          MoveJ speed 100 deg/s, acceleration 80 deg/s^2 (useActiveTCP=true) feature=FRM_Reference
            Waypoint Variable (Variable): motionParameters(blendRadius=0.02); variable=PSE_A
        MoveL speed 400 mm/s, acceleration 500 mm/s^2 (useActiveTCP=true) feature=FRM_Reference
          Waypoint Variable (Variable): motionParameters(jointSpeed=1.047198 jointAcceleration=1.396263 cartesianSpeed=0.09 cartesianAcceleration=0.05); variable=PSE_T
          'ADD OPEN GRIPPER'
          URCap Gripper (Robotiq_Grippers, Robotiq Inc.) dataModel(position=78.82352941176471, force=11.0, speed=0.0, positionInDouble=78.82352941176471, forceInDouble=11.0, speedInDouble=0.0, slaveIds=[9], blocking=true)
          Waypoint Variable (Variable): motionParameters(jointSpeed=1.047198 jointAcceleration=1.396263 cartesianSpeed=0.09 cartesianAcceleration=0.05); variable=PSE_T_H
          URCap Gripper (Robotiq_Grippers, Robotiq Inc.) dataModel(position=24.705882352941178, force=11.0, speed=0.0, positionInDouble=24.705882352941178, forceInDouble=11.0, speedInDouble=0.0, slaveIds=[9], blocking=true)
          Waypoint Variable (Variable): variable=PSE_R
    Case (caseValue=7)
      Folder Load [hidden by the author, left out]
    Case (caseValue=8)
      Folder Unload [hidden by the author, left out]
    Case (caseValue=11)
      Folder Place without opening gripper
        Action_Info := "place object without gripper opening"
        SuppressedNode
          Script: do_transition(pose_trans(FRM_Reference, PSE_T), keep_rxry=OBJ_Picked)
        Script: movel(FRM_Container_S, a=0.025, v=0.015, r=0.00001)
        Folder EXTT
          Switch expression=JIG
            Case (caseValue=1)
              Folder 3FG
                If OBJ_Picked
                  Set DigitalOutput pin=GRP_3F_Open; digitalValue=1
        If PSE_A_H≠PSE_Z
          If JNT_Q≠JNT_Z
            Script: movej(get_inverse_kin(pose_trans(FRM_Reference, PSE_A_H), qnear=JNT_Q), r=0.050)
          Else 
            Script: movej(pose_trans(FRM_Reference, PSE_A_H), r=0.050)
        If PSE_A≠PSE_Z
          If JNT_Q≠JNT_Z
            Script: movej(get_inverse_kin(pose_trans(FRM_Reference, PSE_A), qnear=JNT_Q), r=0.020)
          Else 
            Script: movej(pose_trans(FRM_Reference, PSE_A), r=0.020)
        MoveL speed 400 mm/s, acceleration 500 mm/s^2 (useActiveTCP=true) feature=FRM_Reference
          If PSE_T_H≠PSE_Z
            Waypoint Variable (Variable): motionParameters(blendRadius=0.01); variable=PSE_T_H
          Waypoint Variable (Variable): motionParameters(jointSpeed=1.047198 jointAcceleration=1.396263 cartesianSpeed=0.09 cartesianAcceleration=0.05); variable=PSE_T
            Until TOOL_CONTACT_DETECTION (allowActions=false retraction=NONE decelerationAcceleration=0.5 decelerationAngularAcceleration=34.906585)
          Force Frame feature=FRM_Reference; selection=[1, 1, 1, 0, 0, 0]; wrench=[0, 0, 0, 0, 0, 0]; limitsForce=[0.1, 0.1, 0.01, 1.047198, 1.047198, 1.047198]; limitsMotion=[0.1, 0.1, 0.1, 0.349066, 0.349066, 0.349066]
            Waypoint Variable (Variable): motionParameters(jointSpeed=1.047198 jointAcceleration=1.396263 cartesianSpeed=0.07 cartesianAcceleration=0.04); variable=PSE_T
          Folder EXTT
            Switch expression=JIG
              Case (caseValue=1)
                Folder 3FG
                  If OBJ_Picked
                    Set DigitalOutput pin=GRP_3F_Open; digitalValue=0
                    Wait Sleep waitTime=0.2
          Folder EOAT
            ''
    Case (caseValue=12)
      Folder Decap
        Action_Info := "decapping"
        Set DigitalOutput pin=GRP_3F_Enable; digitalValue=1
        Set DigitalOutput pin=GRP_3F_Decap; digitalValue=1
        Force Simple feature=Joint_6_name; selection=[0, 0, 1, 0, 0, 0]; wrench=[0, 0, 5, 0, 0, 0]; limitsForce=[0.15, 0.15, 0.15, 1.047198, 1.047198, 1.047198]; limitsMotion=[0.1, 0.1, 0.1, 0.349066, 0.349066, 0.349066]
          Script: check_decapping(offset=0.015, timeout=5, abort=CMD_Hold)
        Set DigitalOutput pin=GRP_3F_Decap; digitalValue=0
        Set DigitalOutput pin=GRP_3F_Enable; digitalValue=0
        MoveL speed 150 mm/s, acceleration 800 mm/s^2 (useActiveTCP=true) feature=FRM_Reference
          Waypoint Variable (Variable): variable=PSE_R
    Case (caseValue=13)
      Timer (action=Reset) variable(name=TMR_Barcode)
      Folder Read [hidden by the author, left out]
    Case (caseValue=15)
      Folder Detect
        Action_Info := "detect"
    Case (caseValue=30)
      Folder Shake
        Action_Info := "shake"
        Script: do_transition(pose_trans(FRM_Reference, PSE_T), keep_rxry=OBJ_Picked)
        If PSE_A_H≠PSE_Z
          If JNT_Q≠JNT_Z
            Script: movej(get_inverse_kin(pose_trans(FRM_Reference, PSE_A_H), qnear=JNT_Q), r=0.050)
          Else 
            Script: movej(pose_trans(FRM_Reference, PSE_A_H), r=0.050)
        If PSE_A≠PSE_Z
          If JNT_Q≠JNT_Z
            Script: movej(get_inverse_kin(pose_trans(FRM_Reference, PSE_A), qnear=JNT_Q), r=0.020)
          Else 
            Script: movej(pose_trans(FRM_Reference, PSE_A), r=0.020)
        MoveL speed 400 mm/s, acceleration 500 mm/s^2 (useActiveTCP=true) feature=FRM_Reference
          If PSE_T_H≠PSE_Z
            Waypoint Variable (Variable): motionParameters(blendRadius=0.01); variable=PSE_T_H
          Waypoint Variable (Variable): motionParameters(jointSpeed=1.047198 jointAcceleration=1.396263 cartesianSpeed=0.12 cartesianAcceleration=0.08); variable=PSE_T
          Folder EXTT
            ''
            MoveJ speed 60 deg/s, acceleration 80 deg/s^2 (useActiveTCP=true) feature=Base
              Waypoint Waypoint_6: TCP in base x=8.801 y=-547.927 z=402.697 mm, rx=-0.5899 ry=-0.0072 rz=-0.0613 rad; joints [-69.01, -76.872, -104.694, -56.634, 78.043, -158.781] deg; TCP offset x=0 y=0 z=161 mm, rx=3.1415 ry=0 rz=0 rad
            MoveJ speed 60 deg/s, acceleration 80 deg/s^2 (useActiveTCP=true) feature=Base
              Waypoint Waypoint_18: TCP in base x=-178.372 y=-433.927 z=368.082 mm, rx=-0.0866 ry=0.7047 rz=-0.0079 rad; joints [-72.502, -76.524, -102.817, -99.71, 50.308, -158.785] deg
            MoveJ speed 60 deg/s, acceleration 80 deg/s^2 (useActiveTCP=true) feature=Base
              Waypoint Waypoint_12: TCP in base x=8.801 y=-547.927 z=402.697 mm, rx=-0.5899 ry=-0.0072 rz=-0.0613 rad; joints [-69.01, -76.872, -104.694, -56.634, 78.043, -158.781] deg
            MoveJ speed 60 deg/s, acceleration 80 deg/s^2 (useActiveTCP=true) feature=Base
              Waypoint Waypoint_19: TCP in base x=-178.372 y=-433.927 z=368.082 mm, rx=-0.0866 ry=0.7047 rz=-0.0079 rad; joints [-72.502, -76.524, -102.817, -99.71, 50.308, -158.785] deg
          If PSE_R_H≠PSE_Z
            Waypoint Variable (Variable): motionParameters(blendRadius=0.01); variable=PSE_R
            Waypoint Variable (Variable): variable=PSE_R_H
          Else 
            Waypoint Variable (Variable): variable=PSE_R
    Case (caseValue=31)
      Action_Info := "Pick_Vial"
      Folder Pick_Vial
        URCap Gripper (Robotiq_Grippers, Robotiq Inc.) dataModel(position=0.0, force=27.84313725490196, speed=32.15686274509804, positionInDouble=0.0, forceInDouble=27.84313725490196, speedInDouble=32.15686274509804, slaveIds=[9], blocking=true)
        MoveJ speed 60 deg/s, acceleration 80 deg/s^2 (useActiveTCP=true) feature=Base
          Waypoint Vial_above: motionParameters(jointSpeed=0.436332 jointAcceleration=0.523599 cartesianSpeed=0.25 cartesianAcceleration=1.2 blendRadius=0.05); TCP in base x=17.106 y=-652.093 z=184.921 mm, rx=0 ry=0 rz=1.5641 rad; joints [-76.636, -112.403, -84.029, -73.556, 90.141, -256.27] deg
        MoveL speed 250 mm/s, acceleration 1200 mm/s^2 (useActiveTCP=true) feature=Base
          Waypoint Vial_pick_point: motionParameters(jointSpeed=1.047198 jointAcceleration=1.396263 cartesianSpeed=0.1 cartesianAcceleration=0.5); TCP in base x=17.106 y=-648.923 z=93.308 mm, rx=0 ry=0 rz=1.5641 rad; joints [-76.583, -116.742, -92.083, -61.164, 90.132, -256.177] deg
        URCap Gripper (Robotiq_Grippers, Robotiq Inc.) dataModel(position=100.0, force=32.94117647058823, speed=27.84313725490196, positionInDouble=100.0, forceInDouble=32.94117647058823, speedInDouble=27.84313725490196, slaveIds=[9], blocking=true)
        MoveL speed 250 mm/s, acceleration 1200 mm/s^2 (useActiveTCP=true) feature=Base
          Waypoint Waypoint_20: motionParameters(jointSpeed=1.047198 jointAcceleration=1.396263 cartesianSpeed=0.1 cartesianAcceleration=0.5 blendRadius=0.05); TCP in base x=19.228 y=-648.67 z=184.921 mm, rx=0 ry=0 rz=0.0241 rad; joints [-76.382, -111.96, -84.66, -73.372, 90.146, -167.779] deg
        SafeHome (positionOptionType=SPEED_AND_ACCELERATION speed=1.047198 acceleration=1.396263 nextMotionTime=2)
    Case (caseValue=32)
      decap := False
      Folder decap_Vial
        Set DigitalOutput pin=digital_out[5]; digitalValue=1
        MoveJ speed 60 deg/s, acceleration 80 deg/s^2 (useActiveTCP=true) feature=Base
          Waypoint Waypoint_33: motionParameters(jointSpeed=0.436332 jointAcceleration=0.523599 cartesianSpeed=0.25 cartesianAcceleration=1.2 blendRadius=0); TCP in base x=-32.362 y=-348.336 z=391.476 mm, rx=0 ry=0 rz=-0.0047 rad; joints [-72.819, -68.266, -97.918, -103.808, 90.124, -162.602] deg
        MoveL speed 250 mm/s, acceleration 1200 mm/s^2 (useActiveTCP=true) feature=Base
          Waypoint Vial_3FG_place: motionParameters(jointSpeed=1.047198 jointAcceleration=1.396263 cartesianSpeed=0.1 cartesianAcceleration=0.5); TCP in base x=-31.859 y=-349.403 z=145.301 mm, rx=0 ry=0 rz=0 rad; joints [-72.903, -71.756, -132.514, -65.722, 90.129, -162.805] deg
        Set DigitalOutput pin=digital_out[5]; digitalValue=0
        Wait Sleep waitTime=0.5
        MoveL speed 250 mm/s, acceleration 1200 mm/s^2 (useActiveTCP=true) feature=Base
          Waypoint Waypoint_34: motionParameters(jointSpeed=1.047198 jointAcceleration=1.396263 cartesianSpeed=0.1 cartesianAcceleration=0.5 blendRadius=0.05); TCP in base x=-32.362 y=-348.336 z=391.476 mm, rx=0 ry=0 rz=-0.0047 rad; joints [-72.819, -68.266, -97.918, -103.808, 90.124, -162.602] deg
        MoveJ speed 60 deg/s, acceleration 80 deg/s^2 (useActiveTCP=true) feature=Base
          Waypoint cap_dump: motionParameters(jointSpeed=0.436332 jointAcceleration=0.523599 cartesianSpeed=0.25 cartesianAcceleration=1.2); TCP in base x=-139.169 y=-420.164 z=146.096 mm, rx=0 ry=0 rz=0 rad; joints [-90.79, -86.479, -121, -62.513, 90.12, -180.712] deg
        URCap Gripper (Robotiq_Grippers, Robotiq Inc.) dataModel(position=0.0, force=100.0, speed=100.0, positionInDouble=0.0, forceInDouble=100.0, speedInDouble=100.0, slaveIds=[9], blocking=true)
        MoveJ speed 60 deg/s, acceleration 80 deg/s^2 (useActiveTCP=true) feature=Base
          Waypoint Waypoint_35: motionParameters(jointSpeed=0.436332 jointAcceleration=0.523599 cartesianSpeed=0.25 cartesianAcceleration=1.2 blendRadius=0.05); TCP in base x=-32.362 y=-348.336 z=391.476 mm, rx=0 ry=0 rz=-0.0047 rad; joints [-72.819, -68.266, -97.918, -103.808, 90.124, -162.602] deg
        MoveL speed 250 mm/s, acceleration 1200 mm/s^2 (useActiveTCP=true) feature=Base
          Waypoint Vial_3FG_place: motionParameters(jointSpeed=1.047198 jointAcceleration=1.396263 cartesianSpeed=0.1 cartesianAcceleration=0.5); TCP in base x=-31.859 y=-349.403 z=145.301 mm, rx=0 ry=0 rz=0 rad; joints [-72.903, -71.756, -132.514, -65.722, 90.129, -162.805] deg
        URCap Gripper (Robotiq_Grippers, Robotiq Inc.) dataModel(position=100.0, force=100.0, speed=80.0, positionInDouble=100.0, forceInDouble=100.0, speedInDouble=80.0, slaveIds=[9], blocking=true)
        SuppressedNode
          decap := True
        SuppressedNode
          Script: dynamic_upward_motion(0.015, 7)
        SuppressedNode
          MoveL speed 250 mm/s, acceleration 1200 mm/s^2 (useActiveTCP=true) feature=Joint_6_name
            MoveDirectionNode (selectedDirection=ZPlus toolParams=8.0E-4, 0.001) feature=Base
              Until DISTANCE (allowActions=false deceleration=3 distanceNodeType=STOP) Distance=0.01; motionParameters(blendRadius=0)
        SuppressedNode
          decap := False
        Folder Decap
          Action_Info := "decapping"
          Set DigitalOutput pin=GRP_3F_Enable; digitalValue=1
          Set DigitalOutput pin=GRP_3F_Decap; digitalValue=1
          Force Frame feature=Base; selection=[0, 0, 1, 0, 0, 0]; wrench=[0, 0, 1, 0, 0, 0]; limitsForce=[0.15, 0.15, 0.001, 1.047198, 1.047198, 1.047198]; limitsMotion=[0.1, 0.1, 0.1, 0.349066, 0.349066, 0.349066]
            Script: check_decapping(offset=0.015, timeout=10, abort=CMD_Hold)
          Set DigitalOutput pin=GRP_3F_Decap; digitalValue=0
          Set DigitalOutput pin=GRP_3F_Enable; digitalValue=0
          MoveL speed 250 mm/s, acceleration 1200 mm/s^2 (useActiveTCP=true) feature=Base
            Waypoint Waypoint_36: motionParameters(jointSpeed=1.047198 jointAcceleration=1.396263 cartesianSpeed=0.1 cartesianAcceleration=0.5 blendRadius=0.05); TCP in base x=-32.362 y=-348.336 z=391.476 mm, rx=0 ry=0 rz=-0.0047 rad; joints [-72.819, -68.266, -97.918, -103.808, 90.124, -162.602] deg
        MoveJ speed 60 deg/s, acceleration 80 deg/s^2 (useActiveTCP=true) feature=Base
          Waypoint cap_dump: motionParameters(jointSpeed=0.436332 jointAcceleration=0.523599 cartesianSpeed=0.25 cartesianAcceleration=1.2); TCP in base x=-139.169 y=-420.164 z=146.096 mm, rx=0 ry=0 rz=0 rad; joints [-90.79, -86.479, -121, -62.513, 90.12, -180.712] deg
        URCap Gripper (Robotiq_Grippers, Robotiq Inc.) dataModel(position=0.0, force=100.0, speed=80.0, positionInDouble=0.0, forceInDouble=100.0, speedInDouble=80.0, slaveIds=[9], blocking=true)
        MoveJ speed 60 deg/s, acceleration 80 deg/s^2 (useActiveTCP=true) feature=Base
          Waypoint Waypoint_37: motionParameters(jointSpeed=0.436332 jointAcceleration=0.523599 cartesianSpeed=0.25 cartesianAcceleration=1.2 blendRadius=0.036); TCP in base x=-32.362 y=-348.336 z=391.476 mm, rx=0 ry=0 rz=-0.0047 rad; joints [-72.819, -68.266, -97.918, -103.808, 90.124, -162.602] deg
    Case (caseValue=33)
      Folder Shake and liquid transfer
        MoveL speed 250 mm/s, acceleration 1200 mm/s^2 (useActiveTCP=true) feature=Base
          Waypoint Vial_liq_above: motionParameters(jointSpeed=1.047198 jointAcceleration=1.396263 cartesianSpeed=0.1 cartesianAcceleration=0.5); TCP in base x=-25.304 y=-338.759 z=426.628 mm, rx=-1.3159 ry=0.8 rz=-0.9283 rad; joints [-21.713, -86.8, -129.663, 45.096, -43.028, -184.708] deg
          Waypoint Vial_liq_pick_1: motionParameters(jointSpeed=1.047198 jointAcceleration=1.396263 cartesianSpeed=0.1 cartesianAcceleration=0.5); TCP in base x=-2.66 y=-335.985 z=159.39 mm, rx=-1.1505 ry=0.6732 rz=-1.0106 rad; joints [-20.975, -83.1, -137.831, -114.287, 46.064, -14.375] deg
          Waypoint Vial_liq_pick_2: motionParameters(jointSpeed=1.047198 jointAcceleration=1.396263 cartesianSpeed=0.1 cartesianAcceleration=0.5); TCP in base x=-41.402 y=-356.792 z=125.395 mm, rx=-1.1435 ry=0.6511 rz=-0.8787 rad; joints [-25.36, -82.348, -146.215, -101.788, 37.598, -24.648] deg
          URCap Gripper (Robotiq_Grippers, Robotiq Inc.) dataModel(position=100.0, force=27.84313725490196, speed=32.15686274509804, positionInDouble=100.0, forceInDouble=27.84313725490196, speedInDouble=32.15686274509804, slaveIds=[9], blocking=true)
          Wait Sleep waitTime=1
          Set DigitalOutput pin=digital_out[5]; digitalValue=1
          Wait Sleep waitTime=0.5
          Waypoint Vial_liq_above: motionParameters(jointSpeed=1.047198 jointAcceleration=1.396263 cartesianSpeed=0.05 cartesianAcceleration=0.3 blendRadius=0.05); TCP in base x=-25.304 y=-338.759 z=426.628 mm, rx=-1.3159 ry=0.8 rz=-0.9283 rad; joints [-21.713, -86.8, -129.663, 45.096, -43.028, -184.708] deg
        MoveL speed 250 mm/s, acceleration 1200 mm/s^2 (useActiveTCP=true) feature=Base
          Waypoint Liquid_midway: motionParameters(jointSpeed=1.047198 jointAcceleration=1.396263 cartesianSpeed=0.1 cartesianAcceleration=0.5 blendRadius=0); TCP in base x=57.575 y=-583.082 z=306.415 mm, rx=-1.3517 ry=0.1209 rz=-0.0969 rad; joints [-51.29, -97.606, -136.419, 36.185, 44.156, -168.768] deg
          Loop Counting (count=3) loopVariable(name=Loop_1)
            Waypoint shake_1: motionParameters(jointSpeed=1.047198 jointAcceleration=1.396263 cartesianSpeed=0.5 cartesianAcceleration=2); TCP in base x=57.575 y=-583.085 z=306.423 mm, rx=-1.361 ry=-0.1556 rz=-0.4381 rad; joints [-51.29, -97.606, -136.418, 36.185, 44.156, -145.5] deg
            Waypoint shake_2: motionParameters(jointSpeed=1.047198 jointAcceleration=1.396263 cartesianSpeed=0.5 cartesianAcceleration=2); TCP in base x=57.582 y=-583.091 z=306.44 mm, rx=-1.3088 ry=0.3685 rz=0.2149 rad; joints [-51.29, -97.606, -136.416, 36.185, 44.155, -190] deg
          Waypoint drop_above_1: motionParameters(jointSpeed=1.047198 jointAcceleration=1.396263 cartesianSpeed=0.1 cartesianAcceleration=0.5); TCP in base x=268.235 y=-467.784 z=226.22 mm, rx=-1.0278 ry=-0.4308 rz=1.0046 rad; joints [-53.609, -95.474, -138.959, 24.045, 105.829, -198.245] deg
          Waypoint drop_above_2: motionParameters(jointSpeed=1.047198 jointAcceleration=1.396263 cartesianSpeed=0.1 cartesianAcceleration=0.5); TCP in base x=219.042 y=-470.776 z=133.754 mm, rx=-0.313 ry=-0.3444 rz=1.5006 rad; joints [-60.743, -97.429, -119.175, -41.501, 111.324, -235.78] deg
          Waypoint liq_tran_1: motionParameters(jointSpeed=1.047198 jointAcceleration=1.396263 cartesianSpeed=0.05 cartesianAcceleration=0.5 blendRadius=0.008); TCP in base x=213.068 y=-469.567 z=100.231 mm, rx=0.2519 ry=0.2179 rz=1.5928 rad; joints [-44.631, -104.414, -106.819, -71.743, 78.886, -225.335] deg
          Wait Sleep waitTime=1
          Waypoint drop_above_2: motionParameters(jointSpeed=1.047198 jointAcceleration=1.396263 cartesianSpeed=0.1 cartesianAcceleration=0.5); TCP in base x=219.042 y=-470.776 z=133.754 mm, rx=-0.313 ry=-0.3444 rz=1.5006 rad; joints [-60.743, -97.429, -119.175, -41.501, 111.324, -235.78] deg
          Waypoint Waypoint_21: motionParameters(jointSpeed=1.047198 jointAcceleration=1.396263 cartesianSpeed=0.1 cartesianAcceleration=0.5); TCP in base x=187.119 y=-493.959 z=133.754 mm, rx=-0.313 ry=-0.3444 rz=1.5006 rad; joints [-65.422, -99.182, -116.519, -44.234, 112.218, -240.733] deg
          Waypoint liq_tran_2: motionParameters(jointSpeed=1.047198 jointAcceleration=1.396263 cartesianSpeed=0.05 cartesianAcceleration=0.5); TCP in base x=195.958 y=-493.023 z=100.231 mm, rx=0.1607 ry=0.1098 rz=1.5253 rad; joints [-50.52, -104.533, -106.862, -66.514, 83.832, -227.689] deg
          Wait Sleep waitTime=1
          Waypoint drop_above_2: motionParameters(jointSpeed=1.047198 jointAcceleration=1.396263 cartesianSpeed=0.1 cartesianAcceleration=0.5); TCP in base x=219.042 y=-470.776 z=133.754 mm, rx=-0.313 ry=-0.3444 rz=1.5006 rad; joints [-60.743, -97.429, -119.175, -41.501, 111.324, -235.78] deg
          Waypoint drop_above_1: motionParameters(jointSpeed=1.047198 jointAcceleration=1.396263 cartesianSpeed=0.1 cartesianAcceleration=0.5); TCP in base x=268.235 y=-467.784 z=226.22 mm, rx=-1.0278 ry=-0.4308 rz=1.0046 rad; joints [-53.609, -95.474, -138.959, 24.045, 105.829, -198.245] deg
          Waypoint Liquid_midway: motionParameters(jointSpeed=1.047198 jointAcceleration=1.396263 cartesianSpeed=0.1 cartesianAcceleration=0.5); TCP in base x=57.575 y=-583.082 z=306.415 mm, rx=-1.3517 ry=0.1209 rz=-0.0969 rad; joints [-51.29, -97.606, -136.419, 36.185, 44.156, -168.768] deg
        MoveL speed 250 mm/s, acceleration 1200 mm/s^2 (useActiveTCP=true) feature=Base
          Waypoint Vial_drop_above: motionParameters(jointSpeed=1.047198 jointAcceleration=1.396263 cartesianSpeed=0.1 cartesianAcceleration=0.5); TCP in base x=0.325 y=-648.57 z=221.894 mm, rx=-0.8735 ry=1.1659 rz=-1.4827 rad; joints [-60.601, -137.11, -52.92, -147.418, 45.283, -19.072] deg
          Waypoint Vial_liq_drop: motionParameters(jointSpeed=1.047198 jointAcceleration=1.396263 cartesianSpeed=0.1 cartesianAcceleration=0.5); TCP in base x=1.021 y=-647.66 z=92.916 mm, rx=-0.8348 ry=1.0819 rz=-1.5406 rad; joints [-60.917, -140.075, -64.676, -125.954, 46.582, -22.337] deg
          URCap Gripper (Robotiq_Grippers, Robotiq Inc.) dataModel(position=0.0, force=27.84313725490196, speed=32.15686274509804, positionInDouble=0.0, forceInDouble=27.84313725490196, speedInDouble=32.15686274509804, slaveIds=[9], blocking=true)
          Waypoint Vial_drop_above: motionParameters(jointSpeed=1.047198 jointAcceleration=1.396263 cartesianSpeed=0.1 cartesianAcceleration=0.5); TCP in base x=0.325 y=-648.57 z=221.894 mm, rx=-0.8735 ry=1.1659 rz=-1.4827 rad; joints [-60.601, -137.11, -52.92, -147.418, 45.283, -19.072] deg
    Case (caseValue=34)
      SafeHome (positionOptionType=SPEED_AND_ACCELERATION speed=1.047198 acceleration=1.396263 nextMotionTime=2)
      MoveJ speed 60 deg/s, acceleration 80 deg/s^2 (useActiveTCP=true) feature=Base
        Waypoint Waypoint_9: motionParameters(jointSpeed=0.436332 jointAcceleration=0.523599 cartesianSpeed=0.25 cartesianAcceleration=1.2); TCP in base x=206.301 y=-401.796 z=209.941 mm, rx=0 ry=0 rz=1.5608 rad; joints [-45.627, -84.145, -113.025, -72.821, 90.127, -225.014] deg
      MoveL speed 250 mm/s, acceleration 1200 mm/s^2 (useActiveTCP=true) feature=Base
        Waypoint Waypoint_10: motionParameters(jointSpeed=1.047198 jointAcceleration=1.396263 cartesianSpeed=0.1 cartesianAcceleration=0.5); TCP in base x=200.866 y=-400.818 z=105.073 mm, rx=0 ry=0 rz=1.5608 rad; joints [-46.083, -90.669, -123.933, -55.389, 90.105, -225.416] deg
      URCap Gripper (Robotiq_Grippers, Robotiq Inc.) dataModel(position=100.0, force=27.84313725490196, speed=32.15686274509804, positionInDouble=100.0, forceInDouble=27.84313725490196, speedInDouble=32.15686274509804, slaveIds=[9], blocking=true)
      Wait Sleep waitTime=1
      MoveL speed 250 mm/s, acceleration 1200 mm/s^2 (useActiveTCP=true) feature=Base
        Waypoint Waypoint_11: motionParameters(jointSpeed=1.047198 jointAcceleration=1.396263 cartesianSpeed=0.1 cartesianAcceleration=0.5 blendRadius=0.05); TCP in base x=200.866 y=-400.818 z=325.177 mm, rx=0 ry=0 rz=1.5608 rad; joints [-46.018, -81.306, -98.396, -90.289, 90.129, -225.47] deg
      MoveJ speed 60 deg/s, acceleration 80 deg/s^2 (useActiveTCP=true) feature=Base
        Waypoint Waypoint_7: motionParameters(jointSpeed=0.436332 jointAcceleration=0.523599 cartesianSpeed=0.25 cartesianAcceleration=1.2 blendRadius=0.05); TCP in base x=-615.829 y=233.809 z=300 mm, rx=0.0051 ry=0.0087 rz=-2.1118 rad; joints [-188.832, -110.936, -69.076, -89.912, 89.674, -157.919] deg
      MoveL speed 250 mm/s, acceleration 1200 mm/s^2 (useActiveTCP=true) feature=Base
        Waypoint Waypoint_8: motionParameters(jointSpeed=1.047198 jointAcceleration=1.396263 cartesianSpeed=0.1 cartesianAcceleration=0.5); TCP in base x=-615.829 y=233.809 z=13.91 mm, rx=0.0051 ry=0.0087 rz=-2.1118 rad; joints [-188.874, -123.68, -94.539, -51.707, 89.657, -157.833] deg
      URCap Gripper (Robotiq_Grippers, Robotiq Inc.) dataModel(position=0.0, force=27.84313725490196, speed=32.15686274509804, positionInDouble=0.0, forceInDouble=27.84313725490196, speedInDouble=32.15686274509804, slaveIds=[9], blocking=true)
      MoveJ speed 60 deg/s, acceleration 80 deg/s^2 (useActiveTCP=true) feature=Base
        Waypoint Waypoint_7: motionParameters(jointSpeed=0.436332 jointAcceleration=0.523599 cartesianSpeed=0.25 cartesianAcceleration=1.2); TCP in base x=-615.829 y=233.809 z=300 mm, rx=0.0051 ry=0.0087 rz=-2.1118 rad; joints [-188.832, -110.936, -69.076, -89.912, 89.674, -157.919] deg
      SafeHome (positionOptionType=SPEED_AND_ACCELERATION speed=1.047198 acceleration=1.396263 nextMotionTime=2)
      SuppressedNode
        Folder Decap
          Action_Info := "decapping"
          Set DigitalOutput pin=GRP_3F_Enable; digitalValue=1
          Set DigitalOutput pin=GRP_3F_Decap; digitalValue=1
          Force Frame feature=Base; selection=[0, 0, 1, 0, 0, 0]; wrench=[0, 0, 1, 0, 0, 0]; limitsForce=[0.15, 0.15, 0.001, 1.047198, 1.047198, 1.047198]; limitsMotion=[0.1, 0.1, 0.1, 0.349066, 0.349066, 0.349066]
            Script: check_decapping(offset=0.015, timeout=10, abort=CMD_Hold)
          Set DigitalOutput pin=GRP_3F_Decap; digitalValue=0
          Set DigitalOutput pin=GRP_3F_Enable; digitalValue=0
          MoveL speed 250 mm/s, acceleration 1200 mm/s^2 (useActiveTCP=true) feature=Base
            Waypoint Waypoint_5: motionParameters(jointSpeed=1.047198 jointAcceleration=1.396263 cartesianSpeed=0.1 cartesianAcceleration=0.5 blendRadius=0.05); TCP in base x=-31.859 y=-349.402 z=312.809 mm, rx=0 ry=0 rz=0 rad; joints [-72.832, -66.838, -110.376, -92.778, 90.139, -162.834] deg
          MoveJ speed 60 deg/s, acceleration 80 deg/s^2 (useActiveTCP=true) feature=Base
            Waypoint cap_dump: motionParameters(jointSpeed=0.436332 jointAcceleration=0.523599 cartesianSpeed=0.25 cartesianAcceleration=1.2); TCP in base x=-139.169 y=-420.164 z=146.096 mm, rx=0 ry=0 rz=0 rad; joints [-90.79, -86.479, -121, -62.513, 90.12, -180.712] deg
          URCap Gripper (Robotiq_Grippers, Robotiq Inc.) dataModel(position=0.0, force=100.0, speed=100.0, positionInDouble=0.0, forceInDouble=100.0, speedInDouble=100.0, slaveIds=[9], blocking=true)
          MoveJ speed 60 deg/s, acceleration 80 deg/s^2 (useActiveTCP=true) feature=Base
            Waypoint Waypoint_5: motionParameters(jointSpeed=0.436332 jointAcceleration=0.523599 cartesianSpeed=0.25 cartesianAcceleration=1.2 blendRadius=0.05); TCP in base x=-31.859 y=-349.402 z=312.809 mm, rx=0 ry=0 rz=0 rad; joints [-72.832, -66.838, -110.376, -92.778, 90.139, -162.834] deg
          Set DigitalOutput pin=digital_out[5]; digitalValue=1
    Case (caseValue=35)
      Folder Pick the powder container
        SuppressedNode
          MoveJ speed 60 deg/s, acceleration 80 deg/s^2 (useActiveTCP=true) feature=Base
            Waypoint Variable (Variable): variable(featureName=CAM_LM_Cont_S)
        URCap VISOR Robotic App (SensoPart VISOR Robotic, SensoPart Industriesensorik GmbH) dataModel(visorAppTemplate=1); state(isChildrenLocked=true)
          URCap Easy Pick Setup (SensoPart VISOR Robotic, SensoPart Industriesensorik GmbH) dataModel(visorId=0, visorSetJob=true, visorImageAcqSetup=2, visorDetector=1, visorOffsetSet=true, visorCalibSetNo=7, visorJobName=Container, visorImageAcqSource=2, visorSetupStatus=2, Pose(key=visorImageAcqPose, Position(key=posePosition, Length(key=X value=-0.51041 unit=M), Length(key=Y value=0.417301 unit=M), Length(key=Z value=0.464095 unit=M)), Rotation(key=poseRotation, Angle(key=RX value=0.000026 unit=RAD), Angle(key=RY value=-0.000024 unit=RAD), Angle(key=RZ value=-2.896187 unit=RAD))), Pose(key=visorGripPose, Position(key=posePosition, Length(key=X value=-0.52891 unit=M), Length(key=Y value=0.461593 unit=M), Length(key=Z value=-0.178186 unit=M)), Rotation(key=poseRotation, Angle(key=RX value=-0.279814 unit=RAD), Angle(key=RY value=2.118244 unit=RAD), Angle(key=RZ value=-2.110314 unit=RAD))), Feature(key=visorImageAcqFeature name=cont_img_pose)); state(isChildrenLocked=true)
          URCap Process (SensoPart VISOR Robotic, SensoPart Industriesensorik GmbH) dataModel(Variable(key=visorCounterVar, variable(name=easyPickCount, initializeExpression=0)), Variable(key=visorPartsFoundVar, variable(name=easyPickParts, initializeExpression=0))); state(isChildrenLocked=true)
            URCap Image Acquisition Pose (SensoPart VISOR Robotic, SensoPart Industriesensorik GmbH) state(isChildrenLocked=true)
            URCap Object Detected (SensoPart VISOR Robotic, SensoPart Industriesensorik GmbH) state(isChildrenLocked=true)
              Folder Open Gripper
                URCap Gripper (Robotiq_Grippers, Robotiq Inc.) dataModel(position=0.0, force=30.0, speed=40.0, positionInDouble=0.0, forceInDouble=30.0, speedInDouble=40.0, slaveIds=[9], blocking=true)
                MoveJ speed 60 deg/s, acceleration 80 deg/s^2 (useActiveTCP=true) feature=Base
                  Waypoint Waypoint_13: TCP in base x=-479.451 y=284.141 z=125.27 mm, rx=-0.2768 ry=2.0984 rz=-2.1213 rad; joints [-165.671, -112.009, -127.874, -95.426, 1.192, -23.029] deg
              URCap Approach Pose (SensoPart VISOR Robotic, SensoPart Industriesensorik GmbH) dataModel(visorOffsetZ=-50.0); state(isChildrenLocked=true)
              URCap Target Pose (SensoPart VISOR Robotic, SensoPart Industriesensorik GmbH) state(isChildrenLocked=true)
              Folder Close Gripper
                URCap Gripper (Robotiq_Grippers, Robotiq Inc.) dataModel(position=100.0, force=30.19607843137255, speed=40.0, positionInDouble=100.0, forceInDouble=30.19607843137255, speedInDouble=40.0, slaveIds=[9], blocking=true)
              URCap Exit Pose (SensoPart VISOR Robotic, SensoPart Industriesensorik GmbH) dataModel(visorOffsetZ=-50.0); state(isChildrenLocked=true)
            URCap No Object Detected (SensoPart VISOR Robotic, SensoPart Industriesensorik GmbH) dataModel(Variable(key=visorNoObjCountVar, variable(name=easyPickNoObj, initializeExpression=0)))
              Popup Message (haltProgram=false message=No Container detected inputType=Text)
        MoveJ speed 60 deg/s, acceleration 80 deg/s^2 (useActiveTCP=true) feature=Base
          SuppressedNode
            Waypoint Cont_midwa_1: motionParameters(jointSpeed=1.047198 jointAcceleration=1.396263 cartesianSpeed=0.25 cartesianAcceleration=1.2 blendRadius=0.01); TCP in base x=-462.252 y=294.856 z=204.322 mm, rx=-0.3472 ry=2.0343 rz=-2.0655 rad; joints [-166.773, -128.859, -129.893, 70.604, 5.32, -171.145] deg
          Waypoint Waypoint_70: motionParameters(jointSpeed=0.523599 jointAcceleration=0.698132 cartesianSpeed=0.25 cartesianAcceleration=1.2 blendRadius=0); TCP in base x=-472.821 y=292.44 z=207.418 mm, rx=-0.2598 ry=-2.0535 rz=2.0707 rad; joints [-170.164, -118.699, -96.461, -142.976, 25.725, -0.32] deg
          Waypoint Waypoint_2: motionParameters(jointSpeed=0.523599 jointAcceleration=0.872665 cartesianSpeed=0.25 cartesianAcceleration=1.2 blendRadius=0.05); TCP in base x=-312.961 y=-152.991 z=223.61 mm, rx=-0.7453 ry=-1.7139 rz=1.6733 rad; joints [-134.992, -125.122, -83.555, -151.463, 94.666, 2.49] deg
          Waypoint Waypoint_3: motionParameters(jointSpeed=0.523599 jointAcceleration=0.698132 cartesianSpeed=0.25 cartesianAcceleration=1.2 blendRadius=0.05); TCP in base x=-113.75 y=-390.11 z=317.307 mm, rx=-0.5194 ry=-0.8399 rz=1.7569 rad; joints [-108.345, -98.585, -86.606, -121.699, 124.957, 41.411] deg
        MoveL speed 250 mm/s, acceleration 1200 mm/s^2 (useActiveTCP=true) feature=Base
          Waypoint Waypoint_15: motionParameters(jointSpeed=1.047198 jointAcceleration=1.396263 cartesianSpeed=0.1 cartesianAcceleration=0.5 blendRadius=0.05); TCP in base x=29.144 y=-436.802 z=327.885 mm, rx=-0.5216 ry=-0.6236 rz=1.8627 rad; joints [-89.657, -89.204, -96.411, -97.086, 128.129, 64.023] deg
          Waypoint Waypoint_14: motionParameters(jointSpeed=1.047198 jointAcceleration=1.396263 cartesianSpeed=0.1 cartesianAcceleration=0.3); TCP in base x=68.712 y=-569.42 z=285.215 mm, rx=-0.6792 ry=-0.7121 rz=1.394 rad; joints [-90.137, -103.3, -96.148, -70.007, 141.633, 93.932] deg
          Waypoint Waypoint_4: motionParameters(jointSpeed=1.047198 jointAcceleration=1.396263 cartesianSpeed=0.05 cartesianAcceleration=0.3); TCP in base x=-47.22 y=-557.625 z=136.371 mm, rx=-0.6792 ry=-0.7121 rz=1.394 rad; joints [-101.643, -114.727, -100.71, -68.127, 140.302, 75.797] deg
        URCap Gripper (Robotiq_Grippers, Robotiq Inc.) dataModel(position=0.0, force=30.0, speed=40.0, positionInDouble=0.0, forceInDouble=30.0, speedInDouble=40.0, slaveIds=[9], blocking=true)
        MoveL speed 250 mm/s, acceleration 1200 mm/s^2 (useActiveTCP=true) feature=Base
          Waypoint Waypoint_25: motionParameters(jointSpeed=1.047198 jointAcceleration=1.396263 cartesianSpeed=0.1 cartesianAcceleration=0.3); TCP in base x=65.436 y=-569.388 z=287.821 mm, rx=-0.6792 ry=-0.7121 rz=1.394 rad; joints [-90.466, -103.248, -95.699, -70.925, 141.635, 93.398] deg
          Waypoint Waypoint_15: motionParameters(jointSpeed=1.047198 jointAcceleration=1.396263 cartesianSpeed=0.1 cartesianAcceleration=0.5 blendRadius=0.05); TCP in base x=29.144 y=-436.802 z=327.885 mm, rx=-0.5216 ry=-0.6236 rz=1.8627 rad; joints [-89.657, -89.204, -96.411, -97.086, 128.129, 64.023] deg
        SafeHome (positionOptionType=SPEED_AND_ACCELERATION speed=1.047198 acceleration=1.396263 nextMotionTime=2)
        SuppressedNode
          MoveJ speed 60 deg/s, acceleration 80 deg/s^2 (useActiveTCP=true) feature=Base
            Waypoint Container_midwa: motionParameters(blendRadius=0.05); TCP in base x=-379.239 y=-127.191 z=300 mm, rx=0 ry=0 rz=-1.2472 rad; joints [-141.945, -74.312, -107.466, -88.214, 90.137, -160.485] deg
        SuppressedNode
          URCap VISOR Robotic App (SensoPart VISOR Robotic, SensoPart Industriesensorik GmbH) dataModel(visorAppTemplate=1); state(isChildrenLocked=true)
            URCap Easy Pick Setup (SensoPart VISOR Robotic, SensoPart Industriesensorik GmbH) dataModel(visorId=0, visorSetJob=true, visorJobName=Target_container, visorImageAcqSetup=2, visorCalibSetNo=7, visorImageAcqSource=0, visorDetector=1, visorOffsetSet=true, visorSetupStatus=3, Pose(key=visorGripPose, Position(key=posePosition, Length(key=X value=-0.43018 unit=M), Length(key=Y value=0.500077 unit=M), Length(key=Z value=-0.155571 unit=M)), Rotation(key=poseRotation, Angle(key=RX value=0.000011 unit=RAD), Angle(key=RY value=0.000015 unit=RAD), Angle(key=RZ value=-2.896111 unit=RAD))), Pose(key=visorImageAcqPose, Position(key=posePosition, Length(key=X value=-0.391157 unit=M), Length(key=Y value=0.420635 unit=M), Length(key=Z value=0.411587 unit=M)), Rotation(key=poseRotation, Angle(key=RX value=-0.000006 unit=RAD), Angle(key=RY value=-0.000024 unit=RAD), Angle(key=RZ value=-2.896146 unit=RAD)))); state(isChildrenLocked=true)
            URCap Process (SensoPart VISOR Robotic, SensoPart Industriesensorik GmbH) dataModel(Variable(key=visorCounterVar, variable(name=easyPickCount_1, initializeExpression=0)), Variable(key=visorPartsFoundVar, variable(name=easyPickParts_1, initializeExpression=0))); state(isChildrenLocked=true)
              URCap Image Acquisition Pose (SensoPart VISOR Robotic, SensoPart Industriesensorik GmbH) state(isChildrenLocked=true)
              URCap Object Detected (SensoPart VISOR Robotic, SensoPart Industriesensorik GmbH) state(isChildrenLocked=true)
                Folder Open Gripper
                  URCap Gripper (Robotiq_Grippers, Robotiq Inc.) dataModel(position=0.0, force=30.0, speed=40.0, positionInDouble=0.0, forceInDouble=30.0, speedInDouble=40.0, slaveIds=[9], blocking=true)
                URCap Approach Pose (SensoPart VISOR Robotic, SensoPart Industriesensorik GmbH) dataModel(visorOffsetZ=-50.0); state(isChildrenLocked=true)
                URCap Target Pose (SensoPart VISOR Robotic, SensoPart Industriesensorik GmbH) state(isChildrenLocked=true)
                Folder Close Gripper
                  URCap Gripper (Robotiq_Grippers, Robotiq Inc.) dataModel(position=100.0, force=30.19607843137255, speed=40.0, positionInDouble=100.0, forceInDouble=30.19607843137255, speedInDouble=40.0, slaveIds=[9], blocking=true)
                URCap Exit Pose (SensoPart VISOR Robotic, SensoPart Industriesensorik GmbH) dataModel(visorOffsetZ=-50.0); state(isChildrenLocked=true)
              URCap No Object Detected (SensoPart VISOR Robotic, SensoPart Industriesensorik GmbH) dataModel(Variable(key=visorNoObjCountVar, variable(name=easyPickNoObj_1, initializeExpression=0)))
                Popup Message (haltProgram=false message=No Target container is detected inputType=Text)
        SuppressedNode
          MoveJ speed 60 deg/s, acceleration 80 deg/s^2 (useActiveTCP=true) feature=Base
            Waypoint Waypoint_16: motionParameters(jointSpeed=0.698132 jointAcceleration=0.872665 cartesianSpeed=0.25 cartesianAcceleration=1.2); TCP in base x=-389.004 y=141.378 z=266.753 mm, rx=0.0001 ry=-0.0001 rz=-2.8961 rad; joints [-181.152, -76.776, -110.541, -82.676, 90.144, -105.201] deg
            Waypoint Waypoint_17: motionParameters(jointSpeed=0.698132 jointAcceleration=0.872665 cartesianSpeed=0.25 cartesianAcceleration=1.2); TCP in base x=-35.034 y=-360.271 z=346.67 mm, rx=0.0001 ry=0 rz=-1.4195 rad; joints [-73.886, -68.929, -104.178, -96.885, 90.142, -82.58] deg
        SuppressedNode
          Set DigitalOutput pin=digital_out[5]; digitalValue=1
        SuppressedNode
          MoveL speed 250 mm/s, acceleration 1200 mm/s^2 (useActiveTCP=true) feature=Base
            Waypoint Waypoint_22: motionParameters(jointSpeed=1.047198 jointAcceleration=1.396263 cartesianSpeed=0.1 cartesianAcceleration=0.5); TCP in base x=-31.771 y=-348.512 z=220.918 mm, rx=0.0001 ry=0 rz=-1.1964 rad; joints [-72.82, -67.691, -123.366, -78.936, 90.15, -94.217] deg
            Waypoint Waypoint_23: motionParameters(jointSpeed=1.047198 jointAcceleration=1.396263 cartesianSpeed=0.05 cartesianAcceleration=0.3); TCP in base x=-31.891 y=-348.193 z=178.714 mm, rx=0.0001 ry=0 rz=-1.1964 rad; joints [-72.841, -69.405, -128.724, -71.864, 90.145, -94.213] deg
        SuppressedNode
          Set DigitalOutput pin=digital_out[5]; digitalValue=0
        SuppressedNode
          Wait Sleep waitTime=1
        SuppressedNode
          URCap Gripper (Robotiq_Grippers, Robotiq Inc.) dataModel(position=0.0, force=30.19607843137255, speed=40.0, positionInDouble=0.0, forceInDouble=30.19607843137255, speedInDouble=40.0, slaveIds=[9], blocking=true)
        SuppressedNode
          MoveL speed 250 mm/s, acceleration 1200 mm/s^2 (useActiveTCP=true) feature=Base
            Waypoint Waypoint_24: motionParameters(jointSpeed=1.047198 jointAcceleration=1.396263 cartesianSpeed=0.05 cartesianAcceleration=0.3); TCP in base x=-31.773 y=-348.52 z=270.997 mm, rx=0.0001 ry=0 rz=-1.1964 rad; joints [-72.799, -66.725, -116.549, -86.72, 90.151, -94.226] deg
        SuppressedNode
          SafeHome (positionOptionType=SPEED_AND_ACCELERATION speed=1.047198 acceleration=1.396263 nextMotionTime=2)
    Case (caseValue=36)
      SuppressedNode
        MoveL speed 250 mm/s, acceleration 1200 mm/s^2 (useActiveTCP=true) feature=Base
          SuppressedNode
            Waypoint Waypoint_26: TCP in base x=-30.182 y=-347.336 z=210.998 mm, rx=0 ry=0 rz=0 rad; joints [-72.486, -67.792, -124.787, -77.413, 90.141, -162.427] deg
      SuppressedNode
        URCap Gripper (Robotiq_Grippers, Robotiq Inc.) dataModel(position=100.0, force=30.19607843137255, speed=40.0, positionInDouble=100.0, forceInDouble=30.19607843137255, speedInDouble=40.0, slaveIds=[9], blocking=true)
      Folder Decap
        SuppressedNode
          Action_Info := "decapping"
        SuppressedNode
          Set DigitalOutput pin=GRP_3F_Enable; digitalValue=1
        SuppressedNode
          Set DigitalOutput pin=GRP_3F_Decap; digitalValue=1
        SuppressedNode
          Force Frame feature=Base; selection=[0, 0, 1, 0, 0, 0]; wrench=[0, 0, 1, 0, 0, 0]; limitsForce=[0.15, 0.15, 0.001, 1.047198, 1.047198, 1.047198]; limitsMotion=[0.1, 0.1, 0.1, 0.349066, 0.349066, 0.349066]
            Script: check_decapping(offset=0.015, timeout=12, abort=CMD_Hold)
        SuppressedNode
          Set DigitalOutput pin=GRP_3F_Decap; digitalValue=0
        SuppressedNode
          Set DigitalOutput pin=GRP_3F_Enable; digitalValue=0
        SuppressedNode
          MoveL speed 250 mm/s, acceleration 1200 mm/s^2 (useActiveTCP=true) feature=Base
            Waypoint Waypoint_27: motionParameters(jointSpeed=1.047198 jointAcceleration=1.396263 cartesianSpeed=0.1 cartesianAcceleration=0.5 blendRadius=0.05); TCP in base x=-30.361 y=-347.415 z=279.539 mm, rx=0 ry=0 rz=-0.0004 rad; joints [-72.488, -66.465, -115.449, -88.079, 90.139, -162.449] deg
            Waypoint Waypoint_28: motionParameters(jointSpeed=1.047198 jointAcceleration=1.396263 cartesianSpeed=0.1 cartesianAcceleration=0.5 blendRadius=0.05); TCP in base x=-154.725 y=-473.257 z=246.189 mm, rx=0 ry=0 rz=-0.0004 rad; joints [-92.526, -89.454, -102.579, -77.959, 90.132, -182.495] deg
            Waypoint Waypoint_29: motionParameters(jointSpeed=1.047198 jointAcceleration=1.396263 cartesianSpeed=0.1 cartesianAcceleration=0.3); TCP in base x=-145.695 y=-485.909 z=46.677 mm, rx=0 ry=0 rz=-0.0004 rad; joints [-91.444, -104.036, -119.144, -46.812, 90.094, -181.324] deg
        SuppressedNode
          URCap Gripper (Robotiq_Grippers, Robotiq Inc.) dataModel(position=61.24306326304106, force=30.19607843137255, speed=40.0, positionInDouble=61.24306326304106, forceInDouble=30.19607843137255, speedInDouble=40.0, slaveIds=[9], blocking=true)
        SuppressedNode
          MoveL speed 250 mm/s, acceleration 1200 mm/s^2 (useActiveTCP=true) feature=Base
            Waypoint Waypoint_38: motionParameters(jointSpeed=1.047198 jointAcceleration=1.396263 cartesianSpeed=0.1 cartesianAcceleration=0.5 blendRadius=0.05); TCP in base x=-145.695 y=-485.909 z=261.43 mm, rx=0 ry=0 rz=-0.0004 rad; joints [-91.4, -90.37, -99.399, -80.223, 90.132, -181.38] deg
            URCap Gripper (Robotiq_Grippers, Robotiq Inc.) dataModel(position=0.0, force=30.19607843137255, speed=40.0, positionInDouble=0.0, forceInDouble=30.19607843137255, speedInDouble=40.0, slaveIds=[9], blocking=true)
            Waypoint Waypoint_30: motionParameters(jointSpeed=1.047198 jointAcceleration=1.396263 cartesianSpeed=0.1 cartesianAcceleration=0.5 blendRadius=0.05); TCP in base x=-30.182 y=-347.336 z=265.578 mm, rx=0 ry=0 rz=0 rad; joints [-72.462, -66.558, -117.437, -85.997, 90.142, -162.436] deg
            Waypoint Waypoint_31: motionParameters(jointSpeed=1.047198 jointAcceleration=1.396263 cartesianSpeed=0.1 cartesianAcceleration=0.5); TCP in base x=-30.182 y=-347.336 z=175.833 mm, rx=0 ry=0 rz=0 rad; joints [-72.5, -69.38, -129.182, -71.43, 90.136, -162.42] deg
        SuppressedNode
          URCap Gripper (Robotiq_Grippers, Robotiq Inc.) dataModel(position=79.44506104328524, force=30.19607843137255, speed=40.0, positionInDouble=79.44506104328524, forceInDouble=30.19607843137255, speedInDouble=40.0, slaveIds=[9], blocking=true)
        SuppressedNode
          Wait Sleep waitTime=1
        SuppressedNode
          Set DigitalOutput pin=digital_out[5]; digitalValue=1
        SuppressedNode
          MoveL speed 250 mm/s, acceleration 1200 mm/s^2 (useActiveTCP=true) feature=Base
            Waypoint Waypoint_32: motionParameters(jointSpeed=1.047198 jointAcceleration=1.396263 cartesianSpeed=0.1 cartesianAcceleration=0.5 blendRadius=0.05); TCP in base x=-30.182 y=-347.336 z=316.067 mm, rx=0 ry=0 rz=0 rad; joints [-72.438, -66.521, -110.081, -93.39, 90.138, -162.442] deg
        SuppressedNode
          URCap VISOR Robotic App (SensoPart VISOR Robotic, SensoPart Industriesensorik GmbH) dataModel(visorAppTemplate=1); state(isChildrenLocked=true)
            URCap Easy Pick Setup (SensoPart VISOR Robotic, SensoPart Industriesensorik GmbH) dataModel(visorId=0, visorSetJob=true, visorJobName=Weigh_scale, visorImageAcqSetup=2, visorImageAcqSource=1, visorCalibSetNo=9, visorDetector=1, visorSetupStatus=5, visorOffsetSet=true, Pose(key=visorGripPose, Position(key=posePosition, Length(key=X value=-0.66092 unit=M), Length(key=Y value=-0.026261 unit=M), Length(key=Z value=0.113423 unit=M)), Rotation(key=poseRotation, Angle(key=RX value=0.044036 unit=RAD), Angle(key=RY value=-0.006733 unit=RAD), Angle(key=RZ value=-1.658906 unit=RAD)))); state(isChildrenLocked=true)
            URCap Process (SensoPart VISOR Robotic, SensoPart Industriesensorik GmbH) dataModel(Variable(key=visorCounterVar, variable(name=easyPickCount_2, initializeExpression=0)), Variable(key=visorPartsFoundVar, variable(name=easyPickParts_2, initializeExpression=0))); state(isChildrenLocked=true)
              URCap Image Acquisition Pose (SensoPart VISOR Robotic, SensoPart Industriesensorik GmbH) state(isChildrenLocked=true)
              URCap Object Detected (SensoPart VISOR Robotic, SensoPart Industriesensorik GmbH) state(isChildrenLocked=true)
                Folder Open Gripper
                  Wait NoWait
                URCap Approach Pose (SensoPart VISOR Robotic, SensoPart Industriesensorik GmbH) dataModel(visorOffsetZ=-50.0); state(isChildrenLocked=true)
                URCap Target Pose (SensoPart VISOR Robotic, SensoPart Industriesensorik GmbH) state(isChildrenLocked=true)
                Folder Close Gripper
                  URCap Gripper (Robotiq_Grippers, Robotiq Inc.) dataModel(position=0.0, force=30.19607843137255, speed=40.0, positionInDouble=0.0, forceInDouble=30.19607843137255, speedInDouble=40.0, slaveIds=[9], blocking=true)
                URCap Exit Pose (SensoPart VISOR Robotic, SensoPart Industriesensorik GmbH) dataModel(visorOffsetZ=-100.0); state(isChildrenLocked=true)
              URCap No Object Detected (SensoPart VISOR Robotic, SensoPart Industriesensorik GmbH) dataModel(Variable(key=visorNoObjCountVar, variable(name=easyPickNoObj_2, initializeExpression=0)))
                Popup Message (haltProgram=false message=No weigh scale is detected inputType=Text)
        SuppressedNode
          SafeHome (positionOptionType=SPEED_AND_ACCELERATION speed=1.047198 acceleration=1.396263 nextMotionTime=2)
        MoveJ speed 60 deg/s, acceleration 80 deg/s^2 (useActiveTCP=true) feature=Base
          Waypoint Waypoint_39: TCP in base x=137.772 y=-577.76 z=300 mm, rx=0 ry=0 rz=-1.5944 rad; joints [-63.54, -101.785, -81.001, -87.198, 90.144, -62.245] deg
        MoveL speed 250 mm/s, acceleration 1200 mm/s^2 (useActiveTCP=true) feature=Base
          Waypoint Waypoint_41: motionParameters(jointSpeed=1.047198 jointAcceleration=1.396263 cartesianSpeed=0.1 cartesianAcceleration=0.5); TCP in base x=74.223 y=-565.642 z=234.62 mm, rx=-0.5169 ry=0.5292 rz=-1.5296 rad; joints [-54.985, -107.527, -85.329, -102.066, 60.279, -46.981] deg
          Waypoint Waypoint_40: motionParameters(jointSpeed=1.047198 jointAcceleration=1.396263 cartesianSpeed=0.05 cartesianAcceleration=0.3); TCP in base x=39.988 y=-564.833 z=191.055 mm, rx=-0.7676 ry=0.3431 rz=-2.2413 rad; joints [-57.701, -107.406, -92.471, -93.607, 59.17, -6.639] deg
        URCap Gripper (Robotiq_Grippers, Robotiq Inc.) dataModel(position=100.0, force=20.0, speed=30.0, positionInDouble=100.0, forceInDouble=20.0, speedInDouble=30.0, slaveIds=[9], blocking=true)
        Loop Counting (count=2) loopVariable(name=Loop_2)
          MoveL speed 250 mm/s, acceleration 1200 mm/s^2 (useActiveTCP=true) feature=Base
            Waypoint Waypoint_42: motionParameters(jointSpeed=1.047198 jointAcceleration=1.396263 cartesianSpeed=0.5 cartesianAcceleration=1.2 blendRadius=0); TCP in base x=41.363 y=-564.865 z=192.806 mm, rx=0.2785 ry=0.6241 rz=0.7623 rad; joints [-57.586, -107.397, -92.198, -93.963, 59.209, -186.442] deg
            Waypoint Waypoint_43: TCP in base x=41.363 y=-564.865 z=192.806 mm, rx=0.8543 ry=0.2268 rz=2.453 rad; joints [-57.586, -107.392, -92.206, -93.951, 59.208, -288.609] deg
          URCap Gripper (Robotiq_Grippers, Robotiq Inc.) dataModel(position=24.83906770255271, force=20.0, speed=30.19607843137255, positionInDouble=24.83906770255271, forceInDouble=20.0, speedInDouble=30.19607843137255, slaveIds=[9], blocking=true)
          MoveL speed 250 mm/s, acceleration 1200 mm/s^2 (useActiveTCP=true) feature=Base
            Waypoint Waypoint_44: motionParameters(jointSpeed=1.047198 jointAcceleration=1.396263 cartesianSpeed=0.5 cartesianAcceleration=1.2 blendRadius=0); TCP in base x=40.883 y=-564.854 z=192.194 mm, rx=0.1109 ry=0.6592 rz=0.2757 rad; joints [-57.626, -107.402, -92.291, -93.842, 59.196, -157.494] deg
            Waypoint Waypoint_45: TCP in base x=42.648 y=-564.896 z=194.439 mm, rx=-0.4517 ry=0.5632 rz=-1.3434 rad; joints [-57.484, -107.381, -91.951, -94.273, 59.256, -60.779] deg
          URCap Gripper (Robotiq_Grippers, Robotiq Inc.) dataModel(position=78.43137254901961, force=20.0, speed=30.0, positionInDouble=78.43137254901961, forceInDouble=20.0, speedInDouble=30.0, slaveIds=[9], blocking=true)
        MoveL speed 250 mm/s, acceleration 1200 mm/s^2 (useActiveTCP=true) feature=Base
          Waypoint Waypoint_46: motionParameters(jointSpeed=1.047198 jointAcceleration=1.396263 cartesianSpeed=0.05 cartesianAcceleration=0.3); TCP in base x=99.944 y=-566.244 z=267.343 mm, rx=-0.4517 ry=0.5632 rz=-1.3434 rad; joints [-53.041, -108.287, -79.23, -108.385, 61.102, -56.184] deg
          Waypoint Waypoint_47: motionParameters(jointSpeed=1.047198 jointAcceleration=1.396263 cartesianSpeed=0.1 cartesianAcceleration=0.5 blendRadius=0); TCP in base x=99.944 y=-566.244 z=267.343 mm, rx=-0.1017 ry=0.0587 rz=-1.4579 rad; joints [-63.671, -99.121, -88.981, -82.751, 84.056, -70.038] deg
          Waypoint Waypoint_48: motionParameters(jointSpeed=1.047198 jointAcceleration=1.396263 cartesianSpeed=0.25 cartesianAcceleration=1.2); TCP in base x=-136.183 y=-647.487 z=294.248 mm, rx=-0.1017 ry=0.0587 rz=-1.4579 rad; joints [-87.788, -109.526, -72.49, -86.263, 84.243, -94.331] deg
          Waypoint Waypoint_49: TCP in base x=-159.024 y=-641.021 z=47.692 mm, rx=0 ry=0 rz=-1.4579 rad; joints [-92.238, -121.266, -92.571, -56.15, 90.14, -98.675] deg
        URCap Gripper (Robotiq_Grippers, Robotiq Inc.) dataModel(position=33.9400665926748, force=20.0, speed=30.19607843137255, positionInDouble=33.9400665926748, forceInDouble=20.0, speedInDouble=30.19607843137255, slaveIds=[9], blocking=true)
        MoveL speed 250 mm/s, acceleration 1200 mm/s^2 (useActiveTCP=true) feature=Base
          Waypoint Waypoint_50: TCP in base x=-159.024 y=-641.021 z=291.114 mm, rx=0 ry=0 rz=-1.4579 rad; joints [-92.2, -111.308, -69.838, -88.841, 90.151, -98.75] deg
          SafeHome (positionOptionType=SPEED_AND_ACCELERATION speed=1.047198 acceleration=1.396263 nextMotionTime=2)
    Case (caseValue=37)
      SuppressedNode
        Target_weight :=  (valueSource=Operator message=Enter the Target weight to be dispensed in gm valueType=Float)
      Script: zero_scale()
      SuppressedNode
        URCap VISOR Robotic App (SensoPart VISOR Robotic, SensoPart Industriesensorik GmbH) dataModel(visorAppTemplate=1); state(isChildrenLocked=true)
          URCap Easy Pick Setup (SensoPart VISOR Robotic, SensoPart Industriesensorik GmbH) dataModel(visorId=0, visorSetJob=true, visorImageAcqSetup=2, visorImageAcqSource=1, visorDetector=1, visorOffsetSet=true, visorJobName=Spatula_horizontal, visorSetupStatus=3, visorCalibSetNo=9, Pose(key=visorGripPose, Position(key=posePosition, Length(key=X value=-0.430208 unit=M), Length(key=Y value=0.366458 unit=M), Length(key=Z value=0.299985 unit=M)), Rotation(key=poseRotation, Angle(key=RX value=1.35602 unit=RAD), Angle(key=RY value=-0.160954 unit=RAD), Angle(key=RZ value=2.750948 unit=RAD)))); state(isChildrenLocked=true)
          URCap Process (SensoPart VISOR Robotic, SensoPart Industriesensorik GmbH) dataModel(Variable(key=visorCounterVar, variable(name=easyPickCount_3, initializeExpression=0)), Variable(key=visorPartsFoundVar, variable(name=easyPickParts_3, initializeExpression=0))); state(isChildrenLocked=true)
            URCap Image Acquisition Pose (SensoPart VISOR Robotic, SensoPart Industriesensorik GmbH) state(isChildrenLocked=true)
            URCap Object Detected (SensoPart VISOR Robotic, SensoPart Industriesensorik GmbH) state(isChildrenLocked=true)
              Folder Open Gripper
                URCap Gripper (Robotiq_Grippers, Robotiq Inc.) dataModel(position=43.13725490196078, force=20.0, speed=20.0, positionInDouble=43.13725490196078, forceInDouble=20.0, speedInDouble=20.0, slaveIds=[9], blocking=true)
              URCap Approach Pose (SensoPart VISOR Robotic, SensoPart Industriesensorik GmbH) dataModel(visorOffsetZ=-100.0); state(isChildrenLocked=true)
              URCap Target Pose (SensoPart VISOR Robotic, SensoPart Industriesensorik GmbH) state(isChildrenLocked=true)
              Folder Close Gripper
                URCap Gripper (Robotiq_Grippers, Robotiq Inc.) dataModel(position=100.0, force=20.0, speed=30.19607843137255, positionInDouble=100.0, forceInDouble=20.0, speedInDouble=30.19607843137255, slaveIds=[9], blocking=true)
              URCap Exit Pose (SensoPart VISOR Robotic, SensoPart Industriesensorik GmbH) dataModel(visorToolSpeed=100.0, visorToolAcc=300.0, visorOffsetZ=-200.0); state(isChildrenLocked=true)
            URCap No Object Detected (SensoPart VISOR Robotic, SensoPart Industriesensorik GmbH) dataModel(Variable(key=visorNoObjCountVar, variable(name=easyPickNoObj_3, initializeExpression=0)))
              Popup Message (haltProgram=false message=No spatula is detected inputType=Text)
      SuppressedNode
        MoveL speed 150 mm/s, acceleration 600 mm/s^2 (useActiveTCP=true) feature=Base
          Waypoint Spatula_above: TCP in base x=250.274 y=-257.311 z=422.802 mm, rx=0.0001 ry=-0.0002 rz=3.0658 rad; joints [-23.887, -70.693, -91.695, -107.604, 90.116, 70.385] deg
          Waypoint Spatula_pick: TCP in base x=250.962 y=-257.604 z=233.358 mm, rx=0.0001 ry=-0.0002 rz=3.1149 rad; joints [-23.978, -68.964, -120.765, -80.263, 90.139, 67.596] deg
          URCap Gripper (Robotiq_Grippers, Robotiq Inc.) dataModel(position=100.0, force=30.0, speed=30.0, positionInDouble=100.0, forceInDouble=30.0, speedInDouble=30.0, slaveIds=[9], blocking=true)
          Waypoint Spatula_above: TCP in base x=250.274 y=-257.311 z=422.802 mm, rx=0.0001 ry=-0.0002 rz=3.0658 rad; joints [-23.887, -70.693, -91.695, -107.604, 90.116, 70.385] deg
      URCap VISOR Robotic App (SensoPart VISOR Robotic, SensoPart Industriesensorik GmbH) dataModel(visorAppTemplate=1); state(isChildrenLocked=true)
        URCap Easy Pick Setup (SensoPart VISOR Robotic, SensoPart Industriesensorik GmbH) dataModel(visorId=0, visorSetJob=true, visorImageAcqSetup=2, visorCalibSetNo=9, visorDetector=1, visorOffsetSet=true, visorJobName=Weigh_scale, visorImageAcqSource=2, visorSetupStatus=2, Pose(key=visorGripPose, Position(key=posePosition, Length(key=X value=-0.529609 unit=M), Length(key=Y value=-0.217535 unit=M), Length(key=Z value=0.164929 unit=M)), Rotation(key=poseRotation, Angle(key=RX value=1.812999 unit=RAD), Angle(key=RY value=-0.679367 unit=RAD), Angle(key=RZ value=1.655208 unit=RAD))), Feature(key=visorImageAcqFeature name=cont_img_pose)); state(isChildrenLocked=true)
        URCap Process (SensoPart VISOR Robotic, SensoPart Industriesensorik GmbH) dataModel(Variable(key=visorCounterVar, variable(name=easyPickCount_4, initializeExpression=0)), Variable(key=visorPartsFoundVar, variable(name=easyPickParts_4, initializeExpression=0))); state(isChildrenLocked=true)
          URCap Image Acquisition Pose (SensoPart VISOR Robotic, SensoPart Industriesensorik GmbH) state(isChildrenLocked=true)
          URCap Object Detected (SensoPart VISOR Robotic, SensoPart Industriesensorik GmbH) state(isChildrenLocked=true)
            Folder Open Gripper
              MoveL speed 150 mm/s, acceleration 600 mm/s^2 (useActiveTCP=true) feature=Base
                Weight_value := get_weight()
                URCap Gripper (Robotiq_Grippers, Robotiq Inc.) dataModel(position=0.0, force=30.19607843137255, speed=30.19607843137255, positionInDouble=0.0, forceInDouble=30.19607843137255, speedInDouble=30.19607843137255, slaveIds=[9], blocking=true)
                Waypoint Waypoint_53: motionParameters(blendRadius=0.05); TCP in base x=-50.111 y=-357.608 z=335.881 mm, rx=0.0342 ry=0.0203 rz=-0.2849 rad; joints [-75.987, -70.026, -104.542, -97.668, 89.799, -149.681] deg
                Waypoint Spatula_above: TCP in base x=246.204 y=-251.091 z=422.802 mm, rx=0.0001 ry=-0.0002 rz=3.0658 rad; joints [-23.178, -69.684, -92.315, -107.994, 90.116, 71.093] deg
                Waypoint Spatula_pick: TCP in base x=248.137 y=-254.122 z=229.082 mm, rx=0.0001 ry=-0.0002 rz=3.1149 rad; joints [-23.628, -68.334, -121.776, -79.882, 90.14, 67.949] deg
                URCap Gripper (Robotiq_Grippers, Robotiq Inc.) dataModel(position=100.0, force=30.0, speed=30.0, positionInDouble=100.0, forceInDouble=30.0, speedInDouble=30.0, slaveIds=[9], blocking=true)
                Waypoint Spatula_above: TCP in base x=246.204 y=-251.091 z=422.802 mm, rx=0.0001 ry=-0.0002 rz=3.0658 rad; joints [-23.178, -69.684, -92.315, -107.994, 90.116, 71.093] deg
                Popup Message (haltProgram=false message=Connect the vibration motor inputType=Text)
                Script: tare_scale()
                Waypoint container_start: motionParameters(jointSpeed=1.047198 jointAcceleration=1.396263 cartesianSpeed=0.1 cartesianAcceleration=0.3); TCP in base x=200.65 y=-570.239 z=366.327 mm, rx=1.3605 ry=0.0217 rz=2.6816 rad; joints [-43.946, -125.42, -42.472, -147.901, 58.405, 68.096] deg
                Waypoint container_wp_1: motionParameters(jointSpeed=1.047198 jointAcceleration=1.396263 cartesianSpeed=0.05 cartesianAcceleration=0.3); TCP in base x=170.614 y=-572.151 z=294.509 mm, rx=1.2595 ry=-0.0083 rz=2.7877 rad; joints [-46.577, -118.755, -62.143, -128.361, 58.907, 59.792] deg
                Loop Counting (count=1) loopVariable(name=Loop_9)
                  Waypoint Waypoint_55: motionParameters(jointSpeed=1.047198 jointAcceleration=1.396263 cartesianSpeed=0.07 cartesianAcceleration=0.5); TCP in base x=77.281 y=-567.309 z=212.068 mm, rx=1.2595 ry=-0.0083 rz=2.7877 rad; joints [-52.608, -113.129, -83.31, -109.754, 55.252, 54.186] deg
                    SuppressedNode
                      Until TOOL_CONTACT_DETECTION (allowActions=false retraction=-0.002 decelerationAcceleration=0.2 decelerationAngularAcceleration=34.906585)
                  Waypoint Waypoint_56: motionParameters(jointSpeed=1.047198 jointAcceleration=1.396263 cartesianSpeed=0.05 cartesianAcceleration=0.3); TCP in base x=135.568 y=-570.868 z=245.215 mm, rx=1.4769 ry=-0.0183 rz=2.6796 rad; joints [-47.325, -120.782, -69.397, -128.377, 54.155, 64.498] deg
                  Waypoint Waypoint_74: TCP in base x=164.828 y=-574.638 z=193.751 mm, rx=2.0536 ry=-0.0465 rz=2.2743 rad; joints [-43.873, -140.397, -56.644, -155.146, 50.601, 86.552] deg
                  Set AnalogOutput pin=analog_out[0]; analogValue=3
                  Wait Sleep waitTime=2
                  Set AnalogOutput pin=analog_out[0]; analogValue=0
                SuppressedNode
                  Loop Counting (count=1) loopVariable(name=Loop_10)
                    Waypoint Waypoint_1: motionParameters(jointSpeed=1.047198 jointAcceleration=1.396263 cartesianSpeed=0.4 cartesianAcceleration=1.2); TCP in base x=175.61 y=-574.617 z=223.224 mm, rx=1.7438 ry=-0.031 rz=2.516 rad; joints [-43.942, -131.598, -59.719, -142.336, 52.9, 75.006] deg
                    Waypoint Waypoint_56: motionParameters(jointSpeed=1.047198 jointAcceleration=1.396263 cartesianSpeed=0.05 cartesianAcceleration=0.3); TCP in base x=135.568 y=-570.868 z=245.215 mm, rx=1.4769 ry=-0.0183 rz=2.6796 rad; joints [-47.325, -120.782, -69.397, -128.377, 54.155, 64.498] deg
                Waypoint Waypoint_59: motionParameters(jointSpeed=1.047198 jointAcceleration=1.396263 cartesianSpeed=0.05 cartesianAcceleration=0.3); TCP in base x=272.401 y=-578.183 z=239.561 mm, rx=2.127 ry=0.1139 rz=2.1556 rad; joints [-37.816, -154.733, -25.502, -178.522, 53.445, 96.624] deg
                Waypoint Waypoint_58: motionParameters(jointSpeed=1.047198 jointAcceleration=1.396263 cartesianSpeed=0.05 cartesianAcceleration=0.3); TCP in base x=223.649 y=-578.478 z=276.546 mm, rx=2.1743 ry=-0.0441 rz=2.0587 rad; joints [-41.771, -153.265, -25.455, -184.54, 55.381, 96.631] deg
                MoveJ speed 30 deg/s, acceleration 50 deg/s^2 (useActiveTCP=true) feature=Base
                  Waypoint Waypoint_60: motionParameters(jointSpeed=0.349066 jointAcceleration=0.523599 cartesianSpeed=0.25 cartesianAcceleration=1.2 blendRadius=0.05); TCP in base x=-13.316 y=-544.772 z=383.372 mm, rx=2.2082 ry=0.0375 rz=2.0976 rad; joints [-53.447, -120.321, -68.514, -175.377, 39.556, 98.101] deg
                  Waypoint Waypoint_61: motionParameters(jointSpeed=0.349066 jointAcceleration=0.523599 cartesianSpeed=0.25 cartesianAcceleration=1.2 blendRadius=0.05); TCP in base x=-412.189 y=-356.447 z=383.372 mm, rx=1.7517 ry=-0.74 rz=1.6007 rad; joints [-101.195, -120.321, -68.514, -175.377, 39.556, 98.101] deg
            URCap Approach Pose (SensoPart VISOR Robotic, SensoPart Industriesensorik GmbH) dataModel(visorOffsetZ=-50.0, visorJointSpeed=20.0, visorJointAcc=25.0); state(isChildrenLocked=true)
            URCap Target Pose (SensoPart VISOR Robotic, SensoPart Industriesensorik GmbH) dataModel(visorToolSpeed=50.0, visorToolAcc=100.0); state(isChildrenLocked=true)
            Folder Close Gripper
              dispense_pos := get_actual_tcp_pose()
              MoveL speed 250 mm/s, acceleration 1200 mm/s^2 (useActiveTCP=true) feature=Base
                Start_thread := True
                vib_mot_thread := True
                Wait Sleep waitTime=0.5
                Loop While (checkContinuously=true) expression=Weight_value≤Target_weight and tilt_angle≤-0.40
                  current_error := Target_weight-Weight_value
                  Integral_error := Integral_error+current_error*dt
                  derivative := (current_error-previous_error)/dt
                  tilt_increment := (kp*current_error)+(ki*Integral_error)+(kd*derivative)
                  current_pose := get_actual_tcp_pose()
                  tilt_angle := current_pose[4]
                  tilt_pose := pose_trans(current_pose, p[(tilt_increment/5.3), 0, 0, 0, tilt_increment, 0])
                  Script: movel(tilt_pose, a=0.025, v=0.015, r=0.00001)
                  previous_error := current_error
                Start_thread := False
                SuppressedNode
                  Waypoint Waypoint_64: motionParameters(jointSpeed=1.047198 jointAcceleration=1.396263 cartesianSpeed=0.03 cartesianAcceleration=0.1 blendRadius=0.05); TCP in base x=-542.998 y=-117.021 z=221.977 mm, rx=1.8981 ry=-0.7227 rz=1.5827 rad; joints [-123.845, -120.87, -101.018, -172.406, 14.907, 127.864] deg
                Weight_value := get_weight()
                tilt_angle := -1
                Wait Sleep waitTime=0.5
                vib_mot_thread := False
                MoveL speed 50 mm/s, acceleration 300 mm/s^2 (useActiveTCP=true) feature=Base
                  Waypoint Variable (Variable): motionParameters(jointSpeed=0.436332 jointAcceleration=0.523599 cartesianSpeed=0.05 cartesianAcceleration=0.2); variable=dispense_pos
                Integral_error := 0
                current_error := 0
                previous_error := 0
                Set AnalogOutput pin=analog_out[0]; analogValue=0
            URCap Exit Pose (SensoPart VISOR Robotic, SensoPart Industriesensorik GmbH) dataModel(visorOffsetZ=0.0); state(isChildrenLocked=true)
          URCap No Object Detected (SensoPart VISOR Robotic, SensoPart Industriesensorik GmbH) dataModel(Variable(key=visorNoObjCountVar, variable(name=easyPickNoObj_4, initializeExpression=0)))
            Popup Message (haltProgram=false message=No weigh scale detected inputType=Text)
      Folder powder dispensing
        SuppressedNode
          Target_weight := Target_weight/1000
        Loop While (checkContinuously=false) expression=Weight_value<Target_weight
          MoveL speed 50 mm/s, acceleration 300 mm/s^2 (useActiveTCP=true) feature=Base
            Waypoint Waypoint_75: motionParameters(blendRadius=0.05); TCP in base x=-289.464 y=-270.54 z=342.974 mm, rx=1.97 ry=-0.5594 rz=1.8261 rad; joints [-81.04, -96.392, -107.993, -161.533, 41.848, 95.33] deg
            Waypoint After_disp_1: TCP in base x=234.178 y=-585.611 z=246.647 mm, rx=2.1694 ry=-0.0462 rz=2.0859 rad; joints [-41.467, -155.969, -23.918, -182.388, 55.049, 95.343] deg
            Waypoint After_disp_2: TCP in base x=211.085 y=-585.611 z=185.147 mm, rx=2.1694 ry=-0.0462 rz=2.0859 rad; joints [-42.623, -153.723, -37.417, -171.165, 53.943, 95.401] deg
            Waypoint After_disp_3: TCP in base x=125.935 y=-585.611 z=299.546 mm, rx=0.9596 ry=-0.1344 rz=2.8807 rad; joints [-54.056, -115.535, -63.235, -120.118, 65.773, 48.319] deg
            Loop Counting (count=1) loopVariable(name=Loop_11)
              Waypoint Waypoint_55: motionParameters(jointSpeed=1.047198 jointAcceleration=1.396263 cartesianSpeed=0.07 cartesianAcceleration=0.5); TCP in base x=77.281 y=-567.309 z=212.068 mm, rx=1.2595 ry=-0.0083 rz=2.7877 rad; joints [-52.608, -113.129, -83.31, -109.754, 55.252, 54.186] deg
                SuppressedNode
                  Until TOOL_CONTACT_DETECTION (allowActions=false retraction=0 decelerationAcceleration=0.2 decelerationAngularAcceleration=34.906585)
              Waypoint Waypoint_56: motionParameters(jointSpeed=1.047198 jointAcceleration=1.396263 cartesianSpeed=0.05 cartesianAcceleration=0.3); TCP in base x=135.568 y=-570.868 z=245.215 mm, rx=1.4769 ry=-0.0183 rz=2.6796 rad; joints [-47.325, -120.782, -69.397, -128.377, 54.155, 64.498] deg
              Waypoint Waypoint_74: TCP in base x=164.828 y=-574.638 z=193.751 mm, rx=2.0536 ry=-0.0465 rz=2.2743 rad; joints [-43.873, -140.397, -56.644, -155.146, 50.601, 86.552] deg
              Set AnalogOutput pin=analog_out[0]; analogValue=3
              Wait Sleep waitTime=2
              Set AnalogOutput pin=analog_out[0]; analogValue=0
            Waypoint Waypoint_59: motionParameters(jointSpeed=1.047198 jointAcceleration=1.396263 cartesianSpeed=0.05 cartesianAcceleration=0.3); TCP in base x=272.401 y=-578.183 z=239.561 mm, rx=2.127 ry=0.1139 rz=2.1556 rad; joints [-37.816, -154.733, -25.502, -178.522, 53.445, 96.624] deg
            Waypoint Waypoint_58: motionParameters(jointSpeed=1.047198 jointAcceleration=1.396263 cartesianSpeed=0.05 cartesianAcceleration=0.3); TCP in base x=223.649 y=-578.478 z=276.546 mm, rx=2.1743 ry=-0.0441 rz=2.0587 rad; joints [-41.771, -153.265, -25.455, -184.54, 55.381, 96.631] deg
          MoveJ speed 30 deg/s, acceleration 50 deg/s^2 (useActiveTCP=true) feature=Base
            Waypoint Waypoint_60: motionParameters(jointSpeed=0.349066 jointAcceleration=0.523599 cartesianSpeed=0.25 cartesianAcceleration=1.2 blendRadius=0.05); TCP in base x=-13.316 y=-544.772 z=383.372 mm, rx=2.2082 ry=0.0375 rz=2.0976 rad; joints [-53.447, -120.321, -68.514, -175.377, 39.556, 98.101] deg
            Waypoint Waypoint_61: motionParameters(jointSpeed=0.349066 jointAcceleration=0.523599 cartesianSpeed=0.25 cartesianAcceleration=1.2 blendRadius=0.05); TCP in base x=-412.189 y=-356.447 z=383.372 mm, rx=1.7517 ry=-0.74 rz=1.6007 rad; joints [-101.195, -120.321, -68.514, -175.377, 39.556, 98.101] deg
            Waypoint Waypoint_62: motionParameters(jointSpeed=0.349066 jointAcceleration=0.523599 cartesianSpeed=0.25 cartesianAcceleration=1.2); TCP in base x=-542.659 y=-114.282 z=251.262 mm, rx=1.813 ry=-0.6794 rz=1.6553 rad; joints [-123.661, -111.262, -103.952, -159.22, 12.548, 108.767] deg
          MoveL speed 250 mm/s, acceleration 1200 mm/s^2 (useActiveTCP=true) feature=Base
            Start_thread := True
            Waypoint Variable (Variable): motionParameters(jointSpeed=0.436332 jointAcceleration=0.523599 cartesianSpeed=0.05 cartesianAcceleration=0.2); variable=dispense_pos
            vib_mot_thread := True
            Wait Sleep waitTime=0.5
            Loop While (checkContinuously=true) expression=Weight_value≤Target_weight and tilt_angle≤-0.40
              current_error := Target_weight-Weight_value
              Integral_error := Integral_error+current_error*dt
              derivative := (current_error-previous_error)/dt
              tilt_increment := (kp*current_error)+(ki*Integral_error)+(kd*derivative)
              current_pose := get_actual_tcp_pose()
              tilt_angle := current_pose[4]
              tilt_pose := pose_trans(current_pose, p[(tilt_increment/7), 0, 0, 0, tilt_increment, 0])
              Script: movel(tilt_pose, a=0.025, v=0.015, r=0.00001)
              previous_error := current_error
              Wait Sleep waitTime=0.01
            Start_thread := False
            Set AnalogOutput pin=analog_out[0]; analogValue=0
            vib_mot_thread := False
            SuppressedNode
              Waypoint Waypoint_64: motionParameters(jointSpeed=1.047198 jointAcceleration=1.396263 cartesianSpeed=0.03 cartesianAcceleration=0.1 blendRadius=0.05); TCP in base x=-542.998 y=-117.021 z=221.977 mm, rx=1.8981 ry=-0.7227 rz=1.5827 rad; joints [-123.845, -120.87, -101.018, -172.406, 14.907, 127.864] deg
            Weight_value := get_weight()
            tilt_angle := -1
            Wait Sleep waitTime=0.5
          MoveL speed 50 mm/s, acceleration 300 mm/s^2 (useActiveTCP=true) feature=Base
            Waypoint Variable (Variable): motionParameters(jointSpeed=0.436332 jointAcceleration=0.523599 cartesianSpeed=0.05 cartesianAcceleration=0.2); variable=dispense_pos
          Integral_error := 0
          current_error := 0
          previous_error := 0
        MoveL speed 250 mm/s, acceleration 1200 mm/s^2 (useActiveTCP=true) feature=Base
          Waypoint Waypoint_54: motionParameters(jointSpeed=1.047198 jointAcceleration=1.396263 cartesianSpeed=0.1 cartesianAcceleration=0.3); TCP in base x=-289.932 y=-405.861 z=355.714 mm, rx=2.2477 ry=-0.0682 rz=2.0027 rad; joints [-76.592, -102.006, -101.558, -173.509, 21.644, 109.755] deg
          Waypoint After_disp_1: motionParameters(jointSpeed=1.047198 jointAcceleration=1.396263 cartesianSpeed=0.1 cartesianAcceleration=0.4); TCP in base x=234.178 y=-585.611 z=246.647 mm, rx=2.1694 ry=-0.0462 rz=2.0859 rad; joints [-41.467, -155.969, -23.918, -182.388, 55.049, 95.343] deg
          Waypoint After_disp_2: motionParameters(jointSpeed=1.047198 jointAcceleration=1.396263 cartesianSpeed=0.1 cartesianAcceleration=0.4); TCP in base x=211.085 y=-585.611 z=185.147 mm, rx=2.1694 ry=-0.0462 rz=2.0859 rad; joints [-42.623, -153.723, -37.417, -171.165, 53.943, 95.401] deg
          Waypoint After_disp_3: motionParameters(jointSpeed=1.047198 jointAcceleration=1.396263 cartesianSpeed=0.1 cartesianAcceleration=0.4); TCP in base x=125.935 y=-585.611 z=299.546 mm, rx=0.9596 ry=-0.1344 rz=2.8807 rad; joints [-54.056, -115.535, -63.235, -120.118, 65.773, 48.319] deg
          Set AnalogOutput pin=analog_out[0]; analogValue=3
          Wait Sleep waitTime=2
          Set AnalogOutput pin=analog_out[0]; analogValue=0
          Waypoint After_disp_2: TCP in base x=211.085 y=-585.611 z=185.147 mm, rx=2.1694 ry=-0.0462 rz=2.0859 rad; joints [-42.623, -153.723, -37.417, -171.165, 53.943, 95.401] deg
          Waypoint After_disp_1: motionParameters(jointSpeed=1.047198 jointAcceleration=1.396263 cartesianSpeed=0.1 cartesianAcceleration=0.4); TCP in base x=234.178 y=-585.611 z=246.647 mm, rx=2.1694 ry=-0.0462 rz=2.0859 rad; joints [-41.467, -155.969, -23.918, -182.388, 55.049, 95.343] deg
          Waypoint Waypoint_63: motionParameters(blendRadius=0.05); TCP in base x=101.295 y=-465.376 z=381.756 mm, rx=0.9726 ry=-0.1584 rz=2.8872 rad; joints [-48.863, -99.659, -71.872, -130.079, 68.56, 52.636] deg; TCP offset x=0 y=0 z=161 mm, rx=3.1415 ry=0 rz=0 rad
          Waypoint Start: motionParameters(jointSpeed=1.047198 jointAcceleration=1.396263 cartesianSpeed=0.15 cartesianAcceleration=0.6); TCP in base x=-33.065 y=-365.399 z=389.873 mm, rx=0 ry=0 rz=2.7258 rad; joints [-73.774, -70.638, -96.716, -102.629, 90.121, 40.001] deg; TCP offset x=0 y=0 z=161 mm, rx=3.1415 ry=0 rz=0 rad
          Popup Message (haltProgram=false message=Powder dispensed successfully... inputType=Text)
      SuppressedNode
        URCap VISOR Robotic App (SensoPart VISOR Robotic, SensoPart Industriesensorik GmbH) dataModel(visorAppTemplate=1); state(isChildrenLocked=true)
          URCap Easy Pick Setup (SensoPart VISOR Robotic, SensoPart Industriesensorik GmbH) dataModel(visorId=0, visorSetJob=true, visorJobName=Spatula_horizontal, visorImageAcqSetup=2, visorImageAcqSource=0, visorDetector=1, visorOffsetSet=true, visorSetupStatus=1, Pose(key=visorImageAcqPose, Position(key=posePosition, Length(key=X value=-0.477866 unit=M), Length(key=Y value=0.377208 unit=M), Length(key=Z value=0.48314 unit=M)), Rotation(key=poseRotation, Angle(key=RX value=-0.000072 unit=RAD), Angle(key=RY value=-0.000033 unit=RAD), Angle(key=RZ value=-1.610249 unit=RAD))), Pose(key=visorGripPose, Position(key=posePosition, Length(key=X value=-0.547139 unit=M), Length(key=Y value=0.33515 unit=M), Length(key=Z value=0.041533 unit=M)), Rotation(key=poseRotation, Angle(key=RX value=2.188123 unit=RAD), Angle(key=RY value=-0.020843 unit=RAD), Angle(key=RZ value=2.219811 unit=RAD)))); state(isChildrenLocked=true)
          URCap Process (SensoPart VISOR Robotic, SensoPart Industriesensorik GmbH) dataModel(Variable(key=visorCounterVar, variable(name=easyPickCount_5, initializeExpression=0)), Variable(key=visorPartsFoundVar, variable(name=easyPickParts_5, initializeExpression=0))); state(isChildrenLocked=true)
            URCap Image Acquisition Pose (SensoPart VISOR Robotic, SensoPart Industriesensorik GmbH) state(isChildrenLocked=true)
            URCap Object Detected (SensoPart VISOR Robotic, SensoPart Industriesensorik GmbH) state(isChildrenLocked=true)
              Folder Open Gripper
                URCap Gripper (Robotiq_Grippers, Robotiq Inc.) dataModel(position=43.04106548279689, force=30.0, speed=30.0, positionInDouble=43.04106548279689, forceInDouble=30.0, speedInDouble=30.0, slaveIds=[9], blocking=true)
              URCap Approach Pose (SensoPart VISOR Robotic, SensoPart Industriesensorik GmbH) dataModel(visorOffsetZ=-130.0); state(isChildrenLocked=true)
              URCap Target Pose (SensoPart VISOR Robotic, SensoPart Industriesensorik GmbH) state(isChildrenLocked=true)
              Folder Close Gripper
                URCap Gripper (Robotiq_Grippers, Robotiq Inc.) dataModel(position=100.0, force=30.0, speed=30.0, positionInDouble=100.0, forceInDouble=30.0, speedInDouble=30.0, slaveIds=[9], blocking=true)
              URCap Exit Pose (SensoPart VISOR Robotic, SensoPart Industriesensorik GmbH) dataModel(visorOffsetZ=-170.0); state(isChildrenLocked=true)
            URCap No Object Detected (SensoPart VISOR Robotic, SensoPart Industriesensorik GmbH) dataModel(Variable(key=visorNoObjCountVar, variable(name=easyPickNoObj_5, initializeExpression=0)))
              Popup Message (haltProgram=false message=No Spatula detected inputType=Text)
      SuppressedNode
        MoveJ speed 60 deg/s, acceleration 80 deg/s^2 (useActiveTCP=true) feature=Base
          Waypoint Waypoint_1: motionParameters(jointSpeed=1.047198 jointAcceleration=1.396263 cartesianSpeed=0.1 cartesianAcceleration=0.5 blendRadius=0.05); TCP in base x=175.61 y=-574.617 z=223.224 mm, rx=1.7438 ry=-0.031 rz=2.516 rad; joints [-43.942, -131.598, -59.719, -142.336, 52.9, 75.006] deg
          Waypoint Waypoint_51: motionParameters(jointSpeed=1.047198 jointAcceleration=1.396263 cartesianSpeed=0.1 cartesianAcceleration=0.5 blendRadius=0); TCP in base x=-477.866 y=377.208 z=483.14 mm, rx=-0.0001 ry=0 rz=-1.6102 rad; joints [-205.499, -110.086, -42.439, -117.467, 90.106, -203.428] deg
          Waypoint Waypoint_52: TCP in base x=-42.31 y=-356.333 z=399.894 mm, rx=0 ry=0 rz=-0.1228 rad; joints [-74.871, -69.823, -95.716, -104.453, 90.124, -157.892] deg
      SuppressedNode
        MoveL speed 50 mm/s, acceleration 300 mm/s^2 (useActiveTCP=true) feature=Base
          Waypoint Waypoint_73: motionParameters(jointSpeed=1.047198 jointAcceleration=1.396263 cartesianSpeed=0.05 cartesianAcceleration=0.3); TCP in base x=200.65 y=-570.239 z=330.084 mm, rx=1.3605 ry=0.0217 rz=2.6816 rad; joints [-43.952, -124.342, -49.589, -141.868, 58.423, 68.107] deg
          Waypoint Waypoint_65: motionParameters(jointSpeed=1.047198 jointAcceleration=1.396263 cartesianSpeed=0.05 cartesianAcceleration=0.3); TCP in base x=143.03 y=-569.853 z=275.754 mm, rx=1.2979 ry=0.0264 rz=2.7129 rad; joints [-47.784, -117.454, -67.716, -126.008, 56.917, 63.329] deg
          Loop Counting (count=3) loopVariable(name=Loop_3)
            Waypoint Waypoint_55: motionParameters(jointSpeed=1.047198 jointAcceleration=1.396263 cartesianSpeed=0.05 cartesianAcceleration=0.3); TCP in base x=73.857 y=-577.013 z=221.505 mm, rx=1.2979 ry=0.0264 rz=2.7129 rad; joints [-52.913, -114.774, -80.289, -113.397, 53.656, 58.584] deg
              Until TOOL_CONTACT_DETECTION (allowActions=false retraction=0 decelerationAcceleration=3 decelerationAngularAcceleration=34.906585)
            Waypoint Waypoint_56: motionParameters(jointSpeed=1.047198 jointAcceleration=1.396263 cartesianSpeed=0.05 cartesianAcceleration=0.3); TCP in base x=135.677 y=-579.448 z=242.231 mm, rx=1.5554 ry=0.0154 rz=2.5559 rad; joints [-47.427, -124.812, -65.265, -134.284, 52.841, 72.036] deg
          Loop Counting (count=2) loopVariable(name=Loop_5)
            Waypoint Waypoint_56: motionParameters(jointSpeed=1.047198 jointAcceleration=1.396263 cartesianSpeed=0.05 cartesianAcceleration=0.3); TCP in base x=135.677 y=-579.448 z=242.231 mm, rx=1.5554 ry=0.0154 rz=2.5559 rad; joints [-47.427, -124.812, -65.265, -134.284, 52.841, 72.036] deg
            Waypoint Waypoint_57: motionParameters(jointSpeed=1.047198 jointAcceleration=1.396263 cartesianSpeed=0.5 cartesianAcceleration=1.2); TCP in base x=143.391 y=-581.809 z=226.065 mm, rx=1.6397 ry=0.0079 rz=2.5024 rad; joints [-46.773, -128.399, -63.349, -137.511, 52.317, 75.293] deg
          Waypoint Waypoint_59: motionParameters(jointSpeed=1.047198 jointAcceleration=1.396263 cartesianSpeed=0.05 cartesianAcceleration=0.3); TCP in base x=272.401 y=-578.183 z=239.561 mm, rx=2.127 ry=0.1139 rz=2.1556 rad; joints [-37.816, -154.733, -25.502, -178.522, 53.445, 96.624] deg
          Waypoint Waypoint_58: motionParameters(jointSpeed=1.047198 jointAcceleration=1.396263 cartesianSpeed=0.05 cartesianAcceleration=0.3); TCP in base x=223.649 y=-578.478 z=276.546 mm, rx=2.1743 ry=-0.0441 rz=2.0587 rad; joints [-41.771, -153.265, -25.455, -184.54, 55.381, 96.631] deg
      SuppressedNode
        MoveJ speed 30 deg/s, acceleration 50 deg/s^2 (useActiveTCP=true) feature=Base
          Waypoint Waypoint_60: motionParameters(jointSpeed=0.349066 jointAcceleration=0.523599 cartesianSpeed=0.25 cartesianAcceleration=1.2 blendRadius=0.05); TCP in base x=-13.316 y=-544.772 z=383.372 mm, rx=2.2082 ry=0.0375 rz=2.0976 rad; joints [-53.447, -120.321, -68.514, -175.377, 39.556, 98.101] deg
          Waypoint Waypoint_61: motionParameters(jointSpeed=0.349066 jointAcceleration=0.523599 cartesianSpeed=0.25 cartesianAcceleration=1.2 blendRadius=0.05); TCP in base x=-412.189 y=-356.447 z=383.372 mm, rx=1.7517 ry=-0.74 rz=1.6007 rad; joints [-101.195, -120.321, -68.514, -175.377, 39.556, 98.101] deg
          Waypoint Waypoint_62: motionParameters(jointSpeed=0.349066 jointAcceleration=0.523599 cartesianSpeed=0.25 cartesianAcceleration=1.2); TCP in base x=-542.659 y=-114.282 z=251.262 mm, rx=1.813 ry=-0.6794 rz=1.6553 rad; joints [-123.661, -111.262, -103.952, -159.22, 12.548, 108.767] deg
      SuppressedNode
        MoveL speed 250 mm/s, acceleration 1200 mm/s^2 (useActiveTCP=true) feature=Base
          Waypoint Waypoint_63: motionParameters(jointSpeed=1.047198 jointAcceleration=1.396263 cartesianSpeed=0.05 cartesianAcceleration=0.3); TCP in base x=-532.496 y=-127.81 z=159.342 mm, rx=1.813 ry=-0.6794 rz=1.6553 rad; joints [-121.654, -119.526, -108.357, -144.665, 14.532, 106.823] deg
          Waypoint Waypoint_66: motionParameters(jointSpeed=1.047198 jointAcceleration=1.396263 cartesianSpeed=0.05 cartesianAcceleration=0.3); TCP in base x=-576.035 y=-66.27 z=306.74 mm, rx=0.8621 ry=-0.2554 rz=2.1952 rad; joints [-142.141, -87.685, -107.535, -64.498, 50.077, -8.596] deg
          Waypoint Waypoint_69: motionParameters(jointSpeed=1.047198 jointAcceleration=1.396263 cartesianSpeed=0.05 cartesianAcceleration=0.3); TCP in base x=-581.965 y=-59.291 z=312.082 mm, rx=0.8621 ry=-0.2554 rz=2.1952 rad; joints [-143.275, -88.018, -106.65, -64.116, 50.29, -10.05] deg
          Waypoint Waypoint_71: motionParameters(jointSpeed=1.047198 jointAcceleration=1.396263 cartesianSpeed=0.5 cartesianAcceleration=1.2); TCP in base x=-581.965 y=-59.291 z=290.576 mm, rx=0.8621 ry=-0.2554 rz=2.1952 rad; joints [-143.281, -88.87, -109.094, -60.824, 50.286, -10.043] deg
          Waypoint Waypoint_72: TCP in base x=-581.965 y=-59.291 z=350.142 mm, rx=1.7575 ry=-0.6778 rz=1.6965 rad; joints [-131.863, -101.687, -97.87, -162.913, 4.302, 96.426] deg
      SuppressedNode
        MoveJ speed 60 deg/s, acceleration 80 deg/s^2 (useActiveTCP=true) feature=Base
          Waypoint Waypoint_68: TCP in base x=-333.293 y=-480.744 z=350.142 mm, rx=2.2175 ry=0.1409 rz=2.2091 rad; joints [-82.414, -101.687, -97.87, -162.913, 4.302, 96.426] deg
      SuppressedNode
        Weight_value := get_weight()
    Case (caseValue=38)
      Folder PowderA(M200)
        URCap VISOR Robotic App (SensoPart VISOR Robotic, SensoPart Industriesensorik GmbH) dataModel(visorAppTemplate=1); state(isChildrenLocked=true)
          URCap Easy Pick Setup (SensoPart VISOR Robotic, SensoPart Industriesensorik GmbH) dataModel(visorId=0, visorSetJob=true, visorJobName=PowderA, visorImageAcqSetup=2, visorImageAcqSource=2, visorDetector=1, visorOffsetSet=true, visorSetupStatus=5, Pose(key=visorGripPose, Position(key=posePosition, Length(key=X value=-0.528934 unit=M), Length(key=Y value=0.461578 unit=M), Length(key=Z value=-0.178169 unit=M)), Rotation(key=poseRotation, Angle(key=RX value=-0.279881 unit=RAD), Angle(key=RY value=2.118252 unit=RAD), Angle(key=RZ value=-2.110291 unit=RAD))), Feature(key=visorImageAcqFeature name=FRM_Container_S)); state(isChildrenLocked=true)
          URCap Process (SensoPart VISOR Robotic, SensoPart Industriesensorik GmbH) dataModel(Variable(key=visorCounterVar, variable(name=easyPickCount_6, initializeExpression=0)), Variable(key=visorPartsFoundVar, variable(name=easyPickParts_6, initializeExpression=0))); state(isChildrenLocked=true)
            URCap Image Acquisition Pose (SensoPart VISOR Robotic, SensoPart Industriesensorik GmbH) state(isChildrenLocked=true)
            URCap Object Detected (SensoPart VISOR Robotic, SensoPart Industriesensorik GmbH) state(isChildrenLocked=true)
              Folder Open Gripper
                URCap Gripper (Robotiq_Grippers, Robotiq Inc.) dataModel(position=0.0, force=30.0, speed=30.0, positionInDouble=0.0, forceInDouble=30.0, speedInDouble=30.0, slaveIds=[9], blocking=true)
                MoveJ speed 60 deg/s, acceleration 80 deg/s^2 (useActiveTCP=true) feature=Base
                  Waypoint Waypoint_76: TCP in base x=-479.451 y=284.141 z=125.27 mm, rx=-0.2768 ry=2.0984 rz=-2.1213 rad; joints [-165.671, -112.009, -127.874, -95.426, 1.192, -23.029] deg
              URCap Approach Pose (SensoPart VISOR Robotic, SensoPart Industriesensorik GmbH) dataModel(visorOffsetZ=-50.0); state(isChildrenLocked=true)
              URCap Target Pose (SensoPart VISOR Robotic, SensoPart Industriesensorik GmbH) state(isChildrenLocked=true)
              Folder Close Gripper
                URCap Gripper (Robotiq_Grippers, Robotiq Inc.) dataModel(position=96.86274509803921, force=30.0, speed=30.0, positionInDouble=96.86274509803921, forceInDouble=30.0, speedInDouble=30.0, slaveIds=[9], blocking=true)
              URCap Exit Pose (SensoPart VISOR Robotic, SensoPart Industriesensorik GmbH) dataModel(visorOffsetZ=-50.0); state(isChildrenLocked=true)
            URCap No Object Detected (SensoPart VISOR Robotic, SensoPart Industriesensorik GmbH) dataModel(Variable(key=visorNoObjCountVar, variable(name=easyPickNoObj_6, initializeExpression=0)))
              Popup Message (haltProgram=false message=No Powder container is detected inputType=Text)
  '=========='
  Folder PostSettings [hidden by the author, left out]
